RoboDK station: reto.rdk

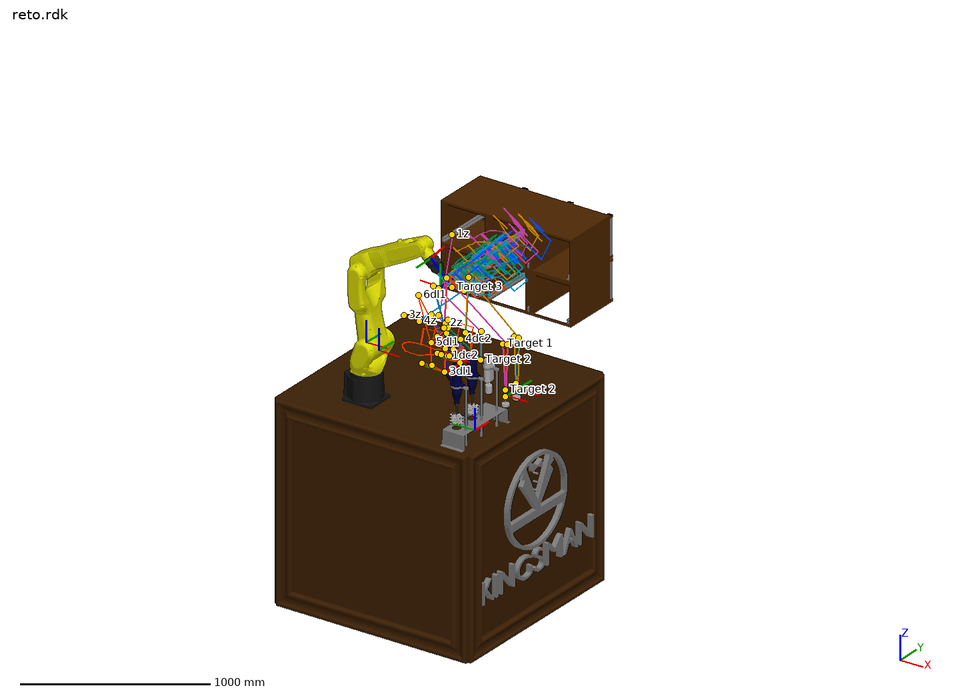
[picture v0: the station drawn from its stored meshes, robots at their saved joint values, targets as dots, program paths as lines]
Station reto (saved by RoboDK 5.5.4). Poses are relative to the parent item; angles as X-Y-Z fixed-axis rotations.
  - frame Fanuc LR Mate 200iD/7L Base at (0, 670, 330) mm
    - robot Fanuc LR Mate 200iD/7L: 6 axes, payload 7 kg, reach 911 mm, repeatability 0.03 mm, weight 27 kg
        modified DH rows (alpha deg, a mm, theta deg, d mm): 0, 0, 0, 330; -90, 50, -90, 0; 0, 440, 0, 0; -90, 35, 0, 420; 90, 0, 0, 0; -90, 0, 0, 80
        base shift (0, 0, -330) mm
        joint limits [-170, -70, -70, -190, -115, -360] to [170, 145, 215, 190, 115, 360]; home [0, 0, 0, 0, 0, 0]; saved at [0, -7.035, 27.253, 0, -70.54, 0]
      - frame RobotiQ 2F-140 Gripper (Mechanism) Base at (0, 0, 0) mm
        - robot RobotiQ 2F-140 Gripper (Mechanism) (model RobotiQ 2F140): 1 axes, payload 5 kg
            joint limits [0] to [140]; home [140]; saved at [30]
          - tool Tool 1, TCP at (0, 0, 190) mm
        - target open (joint target) at (-0.21, -35.16, 190) mm, rotated rx 0 ry -3.02 rz -0.35 deg; joints [30] of RobotiQ 2F-140 Gripper (Mechanism)
        - target close (joint target) at (-114.65, -295.92, 10.81) mm, rotated rx -1.72 ry 2.03 rz 11.69 deg; joints [10] of RobotiQ 2F-140 Gripper (Mechanism)
        - target Target 3 (Cartesian target) at (0, 0, 190) mm; joints [23.986, 137.128, 3.759, 0, 86.241, -156.014] of Fanuc LR Mate 200iD/7L
        - target Target 4 (Cartesian target) at (0, 0, 190) mm; joints [23.986, 137.128, 3.759, 0, 86.241, -156.014] of Fanuc LR Mate 200iD/7L
    - target home (Cartesian target) at (550, 0, 475) mm, rotated rx -180 ry -46.71 rz 0 deg; joints [0, 3.939, 7.691, 0, -50.978, 0] of Fanuc LR Mate 200iD/7L
  - frame rack at (-170, 1590, 240) mm, rotated rx 90 ry 0 rz 180 deg
    - object FullRack (1) at (-810, 360, -320) mm, size 835 x 510 x 385.3 mm, geometry from FullRack (1).STEP
    - target 1z (Cartesian target) at (-358.1, 564.97, -403.2) mm, rotated rx -26.57 ry -40.12 rz 107.86 deg; joints [70, -7.04, 27.25, 0, -70.54, 0] of Fanuc LR Mate 200iD/7L
    - target 2z (Cartesian target) at (-342.39, 58.73, -444.89) mm, rotated rx 2.43 ry -28.49 rz 101.39 deg; joints [48.708, 3.516, -60.085, -111.282, -47, 134.319] of Fanuc LR Mate 200iD/7L
    - target 3z (Cartesian target) at (-104.58, 56.68, -482.72) mm, rotated rx 2.43 ry -28.49 rz 101.39 deg; joints [97.474, -14.415, -55.536, -177.531, -28.246, 164.28] of Fanuc LR Mate 200iD/7L
    - target 4z (Cartesian target) at (-165.76, 16.78, -430.34) mm, rotated rx 2.43 ry -28.49 rz 101.39 deg; joints [82.687, 5.107, -71.647, -159.69, -45.234, 158.787] of Fanuc LR Mate 200iD/7L
    - target 5z (Cartesian target) at (-150, 20, 0) mm, rotated rx 2.43 ry -28.49 rz 101.39 deg; joints [88.603, 43.78, -43.517, 30.239, 18.18, -38.415] of Fanuc LR Mate 200iD/7L
    - target subida charola (Cartesian target) at (-343.88, 69.1, -423.53) mm, rotated rx -21.12 ry -28.57 rz 104.68 deg; joints [68.168, -3.801, -53.905, 12.841, 22.763, -13.527] of Fanuc LR Mate 200iD/7L
  - frame base herramental at (710, 650, 20) mm, rotated rx 0 ry 0 rz 90 deg
    - object Soporte de herramientas at (0, 0, 70) mm, rotated rx 90 ry 0 rz 180 deg, size 443.6 x 340 x 140 mm, geometry from Soporte de herramientas.STEP
  - frame dremel2 at (620, 650, 390) mm, rotated rx 0 ry 0 rz 90 deg
    - target 1dc2 (Cartesian target) at (0.49, 88.9, 17.55) mm, rotated rx -180 ry -61.75 rz -90 deg; joints [89.913, -3.297, -48.984, 180.078, 102.766, 0.058] of Fanuc LR Mate 200iD/7L
    - target 2dc2 (Cartesian target) at (0, 151.76, 13.3) mm, rotated rx -180 ry -61.75 rz -90 deg; joints [-4.961, -25.961, -32.248, 48.26, 5.86, -45.758] of Fanuc LR Mate 200iD/7L
    - target 3dc2 (Cartesian target) at (0, 4.92, 1.2) mm, rotated rx -180 ry -49.6 rz -90 deg; joints [-2.796, -1.172, -33.671, 162.466, 7.084, -160.778] of Fanuc LR Mate 200iD/7L
    - target 4dc2 (Cartesian target) at (0, 0.76, 138.38) mm, rotated rx -180 ry -49.6 rz -90 deg; joints [-2.768, -6.859, -13.429, 175.365, 27.075, -174.076] of Fanuc LR Mate 200iD/7L
    - target 5dc2 (Cartesian target) at (0, 92.68, 148.84) mm, rotated rx -180 ry -44.51 rz -90 deg; joints [-3.386, -17.516, -7.24, 176.175, 38.363, -174.583] of Fanuc LR Mate 200iD/7L
    - target 6dc2 (Cartesian target) at (477.83, 510, 116.81) mm, rotated rx -180 ry -49.6 rz 3.55 deg; joints [64.081, -25.306, -11.026, 143.659, 39.225, -130.203] of Fanuc LR Mate 200iD/7L
  - frame dremel1 at (620, 510.31, 389.97) mm, rotated rx 0 ry 0 rz 90 deg
    - target 1dl1 (Cartesian target) at (0.49, 88.9, 17.55) mm, rotated rx -180 ry -61.75 rz -90 deg; joints [-28.495, -9.165, -37.687, 76.78, 25.575, -60.993] of Fanuc LR Mate 200iD/7L
    - target 2dl1 (Cartesian target) at (0, 151.76, 13.3) mm, rotated rx -180 ry -61.75 rz -90 deg; joints [-34.725, -17.114, -36.143, 84.899, 30.251, -65.939] of Fanuc LR Mate 200iD/7L
    - target 3dl1 (Cartesian target) at (0, 4.92, 1.2) mm, rotated rx -180 ry -49.6 rz -90 deg; joints [-21.306, 2.651, -33.616, 117.955, 18.257, -105.014] of Fanuc LR Mate 200iD/7L
    - target 4dl1 (Cartesian target) at (0, 0.76, 138.38) mm, rotated rx -180 ry -48.03 rz -90 deg; joints [-20.886, -2.493, -13.042, 151.816, 34.141, -141.769] of Fanuc LR Mate 200iD/7L
    - target 5dl1 (Cartesian target) at (0, 92.68, 148.84) mm, rotated rx -180 ry -49.6 rz -90 deg; joints [-26.4, -14.504, -10.508, 146.56, 37.916, -134.648] of Fanuc LR Mate 200iD/7L
    - target 6dl1 (Cartesian target) at (477.83, 510, 116.81) mm, rotated rx -180 ry -55.33 rz 3.55 deg; joints [37.94, -45.517, -1.764, 129.234, 61.201, -109.727] of Fanuc LR Mate 200iD/7L
    - object cepillo1 at (0, -70, -50) mm, rotated rx 90 ry 0 rz 180 deg, size 80 x 351.1 x 124.1 mm, geometry from Dremel con brida.STEP
  - frame bote cera at (140, 586, 355) mm
    - target Target 1 (Cartesian target) at (316.19, 84, 136.54) mm, rotated rx -180 ry -46.71 rz 0 deg; joints [0, -28.492, -10.215, 0, -33.072, 0] of Fanuc LR Mate 200iD/7L
    - target Target 3 (Cartesian target) at (300.65, 202.07, 136.5) mm, rotated rx -180 ry -46.9 rz 15 deg; joints [15, -28.576, -10.266, 0, -32.834, 0] of Fanuc LR Mate 200iD/7L
    - target Target 2 (Cartesian target) at (513.63, 198.92, 10) mm, rotated rx -180 ry -50.56 rz 10.82 deg; joints [9.584, 6.819, -37.897, -31.652, -1.82, 32.424] of Fanuc LR Mate 200iD/7L
    - target Target 4 (Cartesian target) at (516.39, 196.06, 177.59) mm, rotated rx -179.95 ry -49.71 rz 10.96 deg; joints [9.091, -0.877, -13.325, -3.243, -27.022, 4.097] of Fanuc LR Mate 200iD/7L
    - target Target 5 (Cartesian target) at (-35.2, 592.88, 112.91) mm, rotated rx 179.59 ry -46.7 rz 80 deg; joints [77.715, -18.214, -17.774, -2.891, -25.565, 4.172] of Fanuc LR Mate 200iD/7L
  - program open (3 instructions, listed below)
  - program close (3 instructions, listed below)
  - program home (4 instructions, listed below)
  - object mesa at (-1220, 1130, 330) mm, size 1277.5 x 1274.9 x 1205 mm, geometry from mesa.STEP
  - frame zapato at (110, 1270, 40) mm
    - target Target 1 (Cartesian target) at (78.1, -83.2, 764.97) mm, rotated rx -180 ry -46.71 rz 70 deg; joints [70, -7.04, 27.25, 0, -70.54, 0] of Fanuc LR Mate 200iD/7L
    - target Target 2 (Cartesian target) at (48.8, -163.69, 316.74) mm, rotated rx -179.51 ry -45.09 rz 70 deg; joints [69.514, -19.906, -32.534, -3.891, -12.407, 4.144] of Fanuc LR Mate 200iD/7L
    - target Target 3 (Cartesian target) at (51.99, -36.78, 68.56) mm, rotated rx -167.65 ry -61.99 rz 84.86 deg; joints [58.654, 42.845, -90.321, 40.028, 62.94, -6.257] of Fanuc LR Mate 200iD/7L
    - target Target 4 (Cartesian target) at (0, 0, 0) mm, rotated rx -154.66 ry -59.5 rz 70 deg; joints [67.996, 54.587, -97.1, 29.193, 68.847, -10.257] of Fanuc LR Mate 200iD/7L
    - target Target 5 (Cartesian target) at (-12.96, -146.91, 298.71) mm, rotated rx -168.48 ry -59.46 rz 67.92 deg; joints [74.53, -18.6, -45.29, -158.86, -16.3, 156.27] of Fanuc LR Mate 200iD/7L
    - target Target 6 (Cartesian target) at (14.48, -93.65, 48.92) mm, rotated rx -154.66 ry -59.5 rz 70 deg; joints [59.102, 46.97, -102.654, -143.53, -72.674, 174.279] of Fanuc LR Mate 200iD/7L
  - program recoger cepillo cera (10 instructions, listed below)
  - program reset (1 instructions, listed below)
  - program recoger cepillo limpieza (10 instructions, listed below)
  - program recoger cera (9 instructions, listed below)
  - program pick charola (8 instructions, listed below)
  - program c1 recoger (7 instructions, listed below)
  - program c1 entregar (7 instructions, listed below)
  - program poscharolamesa (7 instructions, listed below)
  - program dejar cepillo limpieza (9 instructions, listed below)
  - program dejar cepillo cera (10 instructions, listed below)
  - program dejar  cera (9 instructions, listed below)
  - machining project parribaizq: rotZ(0) | rotX(0)*rotY(0) | onStart | onPathStart | onApproach | onPoint | onRetract | onFinish | SetRPM(%1) | SetTool(%1) | Extruder(%1) | default | default | OutOnMov(%1) | OutOffMov(%1) | onPathFinish | M_RunCode(%1)
  - machining project plateralesizq: rotZ(0) | rotX(0)*rotY(0) | onStart | onPathStart | onApproach | onPoint | onRetract | onFinish | SetRPM(%1) | SetTool(%1) | Extruder(%1) | default | default | OutOnMov(%1) | OutOffMov(%1) | onPathFinish | M_RunCode(%1)
  - program parrizq (66 instructions, listed below)
  - machining project Path3 ajustes: rotZ(0) | rotX(0)*rotY(0) | onStart | onPathStart | onApproach | onPoint | onRetract | onFinish | SetRPM(%1) | SetTool(%1) | Extruder(%1) | default | default | OutOnMov(%1) | OutOffMov(%1) | onPathFinish | M_RunCode(%1)
  - machining project Path4 ajustes: rotZ(0) | rotX(0)*rotY(0) | onStart | onPathStart | onApproach | onPoint | onRetract | onFinish | SetRPM(%1) | SetTool(%1) | Extruder(%1) | default | default | OutOnMov(%1) | OutOffMov(%1) | onPathFinish | M_RunCode(%1)
  - program parrder (59 instructions, listed below)
  - program final (30 instructions, listed below)
  - machining project Path5 ajustes: rotZ(0) | rotX(0)*rotY(0) | onStart | onPathStart | onApproach | onPoint | onRetract | onFinish | SetRPM(%1) | SetTool(%1) | Extruder(%1) | default | default | OutOnMov(%1) | OutOffMov(%1) | onPathFinish | M_RunCode(%1)
  - program cerlatizq (163 instructions, listed below)
  - program platder (154 instructions, listed below)
  - machining project Path6 ajustes: rotZ(0) | rotX(0)*rotY(0) | onStart | onPathStart | onApproach | onPoint | onRetract | onFinish | SetRPM(%1) | SetTool(%1) | Extruder(%1) | default | default | OutOnMov(%1) | OutOffMov(%1) | onPathFinish | M_RunCode(%1)
  - program platizq (163 instructions, listed below)
  - program carribizq (66 instructions, listed below)
  - machining project Path7 ajustes: rotZ(0) | rotX(0)*rotY(0) | onStart | onPathStart | onApproach | onPoint | onRetract | onFinish | SetRPM(%1) | SetTool(%1) | Extruder(%1) | default | default | OutOnMov(%1) | OutOffMov(%1) | onPathFinish | M_RunCode(%1)
  - program cerlatder (154 instructions, listed below)
  - machining project Path8 ajustes: rotZ(0) | rotX(0)*rotY(0) | onStart | onPathStart | onApproach | onPoint | onRetract | onFinish | SetRPM(%1) | SetTool(%1) | Extruder(%1) | default | default | OutOnMov(%1) | OutOffMov(%1) | onPathFinish | M_RunCode(%1)
  - program cerarribder (44 instructions, listed below)
  - machining project Path10 ajustes: rotZ(0) | rotX(0)*rotY(0) | onStart | onPathStart | onApproach | onPoint | onRetract | onFinish | SetRPM(%1) | SetTool(%1) | Extruder(%1) | default | default | OutOnMov(%1) | OutOffMov(%1) | onPathFinish | M_RunCode(%1)
  - program talonder (20 instructions, listed below)
  - frame iman izquierdo at (690, 970, 90) mm, rotated rx 0 ry -0.43 rz 0 deg
    - target Target 1 (Cartesian target) at (-16, -10, 304.12) mm, rotated rx -180 ry -3.01 rz 0 deg; joints [23.726, 34.659, -8.597, 1.235, -78.648, -23.94] of Fanuc LR Mate 200iD/7L
    - target Target 2 (Cartesian target) at (-1.94, -10, 36.88) mm, rotated rx -180 ry -3.01 rz 0 deg; joints [23.284, 48.242, -37.276, 1.554, -49.968, -24.255] of Fanuc LR Mate 200iD/7L
    - target Target 3 (Cartesian target) at (-0.39, -10, 0.32) mm, rotated rx -180 ry 2.75 rz 0 deg; joints [22.488, 53.778, -37.823, -1.092, -54.324, -21.835] of Fanuc LR Mate 200iD/7L
    - target Target 4 (Cartesian target) at (14.23, -10, 304.96) mm, rotated rx -180 ry 2.75 rz 0 deg; joints [22.137, 42.684, -3.214, -0.874, -88.934, -22.104] of Fanuc LR Mate 200iD/7L
    - target Target 5 (Cartesian target) at (-604.68, 318.92, 397.91) mm, rotated rx -178.71 ry 2.21 rz 80.14 deg; joints [82.014, 21.757, -2.792, -0.939, -89.319, -1.878] of Fanuc LR Mate 200iD/7L
    - target Target 6 (Cartesian target) at (-653.05, 360.19, 74.8) mm, rotated rx -178.71 ry 0.13 rz 80.09 deg; joints [86.488, 37.843, -40.739, -1.149, -49.231, -5.645] of Fanuc LR Mate 200iD/7L
  - frame iman derecho at (690, 1070, 90) mm
    - target Target 1 (Cartesian target) at (-16, -10, 304.12) mm, rotated rx -180 ry -3.01 rz 0 deg; joints [30.586, 42.114, -3.765, 1.541, -83.645, -30.722] of Fanuc LR Mate 200iD/7L
    - target Target 2 (Cartesian target) at (-1.94, -10, 36.88) mm, rotated rx -180 ry -3.01 rz 0 deg; joints [30.06, 53.677, -32.189, 1.836, -55.219, -31.073] of Fanuc LR Mate 200iD/7L
    - target Target 3 (Cartesian target) at (-0.39, -0.58, 0.32) mm, rotated rx -180 ry 2.75 rz 0 deg; joints [29.619, 60.126, -31.432, -1.553, -60.966, -28.837] of Fanuc LR Mate 200iD/7L
    - target Target 4 (Cartesian target) at (14.23, -10, 304.96) mm, rotated rx -180 ry 2.75 rz 0 deg; joints [28.537, 52.814, 4.62, -1.322, -97.032, -28.672] of Fanuc LR Mate 200iD/7L
    - target Target 5 (Cartesian target) at (-491.92, 250.35, 416.93) mm, rotated rx -178.68 ry 2.41 rz 72.7 deg; joints [72.54, 30.81, 4.62, -1.32, -97.03, 0] of Fanuc LR Mate 200iD/7L
    - target Target 6 (Cartesian target) at (-525.43, 271.58, 73.13) mm, rotated rx -178.86 ry -1.69 rz 77.54 deg; joints [75.764, 40.036, -38.477, -1.565, -49.877, 2.787] of Fanuc LR Mate 200iD/7L
  - program iman izquierdo (13 instructions, listed below)
  - program iman derecho (13 instructions, listed below)
  - program dejar iman izquierdo (12 instructions, listed below)
  - program dejar iman derecho (12 instructions, listed below)
  - machining project Path10 ajustes: rotZ(0) | rotX(0)*rotY(0) | onStart | onPathStart | onApproach | onPoint | onRetract | onFinish | SetRPM(%1) | SetTool(%1) | Extruder(%1) | default | default | OutOnMov(%1) | OutOffMov(%1) | onPathFinish | M_RunCode(%1)
  - program platizch (163 instructions, listed below)
  - machining project Path11 ajustes: rotZ(0) | rotX(0)*rotY(0) | onStart | onPathStart | onApproach | onPoint | onRetract | onFinish | SetRPM(%1) | SetTool(%1) | Extruder(%1) | default | default | OutOnMov(%1) | OutOffMov(%1) | onPathFinish | M_RunCode(%1)
  - program plaizgr (163 instructions, listed below)
  - machining project Path12 ajustes: rotZ(0) | rotX(0)*rotY(0) | onStart | onPathStart | onApproach | onPoint | onRetract | onFinish | SetRPM(%1) | SetTool(%1) | Extruder(%1) | default | default | OutOnMov(%1) | OutOffMov(%1) | onPathFinish | M_RunCode(%1)
  - program pladerch (154 instructions, listed below)
  - machining project Path13 ajustes: rotZ(0) | rotX(0)*rotY(0) | onStart | onPathStart | onApproach | onPoint | onRetract | onFinish | SetRPM(%1) | SetTool(%1) | Extruder(%1) | default | default | OutOnMov(%1) | OutOffMov(%1) | onPathFinish | M_RunCode(%1)
  - program pladergr (154 instructions, listed below)
  - machining project Path14 ajustes: rotZ(0) | rotX(0)*rotY(0) | onStart | onPathStart | onApproach | onPoint | onRetract | onFinish | SetRPM(%1) | SetTool(%1) | Extruder(%1) | default | default | OutOnMov(%1) | OutOffMov(%1) | onPathFinish | M_RunCode(%1)
  - program arrizch (57 instructions, listed below)
  - machining project Path15 ajustes: rotZ(0) | rotX(0)*rotY(0) | onStart | onPathStart | onApproach | onPoint | onRetract | onFinish | SetRPM(%1) | SetTool(%1) | Extruder(%1) | default | default | OutOnMov(%1) | OutOffMov(%1) | onPathFinish | M_RunCode(%1)
  - program arriderch (52 instructions, listed below)
  - machining project Path16 ajustes: rotZ(0) | rotX(0)*rotY(0) | onStart | onPathStart | onApproach | onPoint | onRetract | onFinish | SetRPM(%1) | SetTool(%1) | Extruder(%1) | default | default | OutOnMov(%1) | OutOffMov(%1) | onPathFinish | M_RunCode(%1)
  - program arridergr (59 instructions, listed below)
  - machining project Path17 ajustes: rotZ(0) | rotX(0)*rotY(0) | onStart | onPathStart | onApproach | onPoint | onRetract | onFinish | SetRPM(%1) | SetTool(%1) | Extruder(%1) | default | default | OutOnMov(%1) | OutOffMov(%1) | onPathFinish | M_RunCode(%1)
  - program arriizqgr (57 instructions, listed below)
  - machining project Path18 ajustes: rotZ(0) | rotX(0)*rotY(0) | onStart | onPathStart | onApproach | onPoint | onRetract | onFinish | SetRPM(%1) | SetTool(%1) | Extruder(%1) | default | default | OutOnMov(%1) | OutOffMov(%1) | onPathFinish | M_RunCode(%1)
  - program cerlaizgr (163 instructions, listed below)
  - machining project Path19 ajustes: rotZ(0) | rotX(0)*rotY(0) | onStart | onPathStart | onApproach | onPoint | onRetract | onFinish | SetRPM(%1) | SetTool(%1) | Extruder(%1) | default | default | OutOnMov(%1) | OutOffMov(%1) | onPathFinish | M_RunCode(%1)
  - program cerladergr (154 instructions, listed below)
  - machining project Path20 ajustes: rotZ(0) | rotX(0)*rotY(0) | onStart | onPathStart | onApproach | onPoint | onRetract | onFinish | SetRPM(%1) | SetTool(%1) | Extruder(%1) | default | default | OutOnMov(%1) | OutOffMov(%1) | onPathFinish | M_RunCode(%1)
  - program ceraariizgr (59 instructions, listed below)
  - machining project Path21 ajustes: rotZ(0) | rotX(0)*rotY(0) | onStart | onPathStart | onApproach | onPoint | onRetract | onFinish | SetRPM(%1) | SetTool(%1) | Extruder(%1) | default | default | OutOnMov(%1) | OutOffMov(%1) | onPathFinish | M_RunCode(%1)
  - program cerarridergr (59 instructions, listed below)
  - machining project Path22 ajustes: rotZ(0) | rotX(0)*rotY(0) | onStart | onPathStart | onApproach | onPoint | onRetract | onFinish | SetRPM(%1) | SetTool(%1) | Extruder(%1) | default | default | OutOnMov(%1) | OutOffMov(%1) | onPathFinish | M_RunCode(%1)
  - program cerlatizqch (163 instructions, listed below)
  - machining project Path23 ajustes: rotZ(0) | rotX(0)*rotY(0) | onStart | onPathStart | onApproach | onPoint | onRetract | onFinish | SetRPM(%1) | SetTool(%1) | Extruder(%1) | default | default | OutOnMov(%1) | OutOffMov(%1) | onPathFinish | M_RunCode(%1)
  - program cerlatderch (154 instructions, listed below)
  - machining project Path25 ajustes: rotZ(0) | rotX(0)*rotY(0) | onStart | onPathStart | onApproach | onPoint | onRetract | onFinish | SetRPM(%1) | SetTool(%1) | Extruder(%1) | default | default | OutOnMov(%1) | OutOffMov(%1) | onPathFinish | M_RunCode(%1)
  - program ceraarribderch (59 instructions, listed below)
  - machining project Path26 ajustes: rotZ(0) | rotX(0)*rotY(0) | onStart | onPathStart | onApproach | onPoint | onRetract | onFinish | SetRPM(%1) | SetTool(%1) | Extruder(%1) | default | default | OutOnMov(%1) | OutOffMov(%1) | onPathFinish | M_RunCode(%1)
  - program ceraarribaizqch (59 instructions, listed below)
  - program final_ch (30 instructions, listed below)
  - program final_gr (30 instructions, listed below)
  - object cepillo2 at (690, 650, 340) mm, rotated rx 90 ry 0 rz -90 deg, size 80 x 351.1 x 124.1 mm, geometry from Dremel con brida.STEP
  - object Iman at (688.21, 960, 126.59) mm, rotated rx 90 ry 0 rz 0 deg, size 45.7 x 91.4 x 45.7 mm, geometry from Iman.STEP
  - object Iman at (688.48, 1060.58, 126.61) mm, size 45.7 x 91.4 x 45.7 mm, geometry from Iman.STEP
  - object Grasa  at (650, 792, 370) mm, size 75 x 201.5 x 85 mm, geometry from Grasa (1).STEP
  - object zapatoconcharola at (-21.13, 1591.46, 262.04) mm, rotated rx 0 ry 0 rz -0.01 deg, size 250 x 350 x 100.5 mm, geometry from zapatoconcharola.STEP
    - object Ruta_IZQ at (-60, 470, 60) mm, rotated rx 0 ry 0 rz -90 deg, geometry from Curva importada
    - object R7 at (-105, 460, 60) mm, rotated rx 0 ry 0 rz -90 deg
    - object Ruta_IZQ_ch at (-60, 390, 60) mm, rotated rx 0 ry 0 rz -90 deg, geometry from Curva importada
    - object R7_ch at (-67.5, 380, 60) mm, rotated rx 0 ry 0 rz -90 deg
    - object Ruta_IZQ_gr at (-50, 550, 80) mm, rotated rx 0 ry 0 rz -90 deg, geometry from Curva importada
    - object R7_gr at (-135, 550, 80) mm, rotated rx 0 ry 0 rz -90 deg
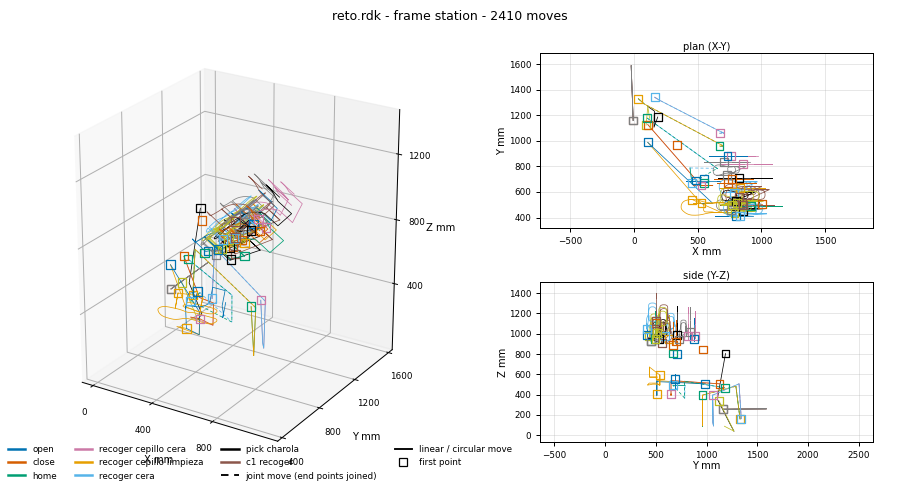
[picture p0: tool path of reto.rdk in frame station, 2410 of 2410 moves have a stored position in this frame; points joined in program order, loops and branches not executed]

--- program open (robot RobotiQ 2F-140 Gripper (Mechanism)) ---
  Est. Ref.: RobotiQ 2F-140 Gripper (Mechanism) Base
  Est. herr: Tool 1
  MoveJ (open)

--- program close (robot RobotiQ 2F-140 Gripper (Mechanism)) ---
  Est. Ref.: RobotiQ 2F-140 Gripper (Mechanism) Base
  Est. herr: Tool 1
  MoveJ (close)

--- program home (robot Fanuc LR Mate 200iD/7L) ---
  Est. Ref.: Fanuc LR Mate 200iD/7L Base
  MoveJ (home)
  Llamar open
  Separar de Tool 1

--- program recoger cepillo cera (robot Fanuc LR Mate 200iD/7L) ---
  Est. Ref.: dremel2
  Est. herr: Tool 1
  MoveL (1dc2)
  MoveL (Target 2) -> target 2dc2
  MoveL (Target 3) -> target 3dc2
  Llamar close
  Adjuntar a Tool 1
  MoveL (Target 4) -> target 4dc2
  MoveL (Target 5) -> target 5dc2
  MoveL (6dc2)

--- program reset (robot Fanuc LR Mate 200iD/7L) ---
  Reemplazar objetos

--- program recoger cepillo limpieza (robot Fanuc LR Mate 200iD/7L) ---
  Est. Ref.: dremel1
  Est. herr: Tool 1
  MoveL (1dl1)
  MoveL (2dl1)
  MoveL (3dl1)
  Adjuntar a Tool 1
  Llamar close
  MoveL (4dl1)
  MoveL (5dl1)
  MoveL (6dl1)

--- program recoger cera (robot Fanuc LR Mate 200iD/7L) ---
  Est. Ref.: bote cera
  Est. herr: Tool 1
  MoveJ (Target 1)
  MoveL (Target 3)
  MoveJ (Target 2)
  Llamar close
  Adjuntar a Tool 1
  MoveJ (Target 4)
  MoveL (Target 5)

--- program pick charola (robot Fanuc LR Mate 200iD/7L) ---
  Est. Ref.: zapato
  Est. herr: Tool 1
  MoveJ (Target 1)
  MoveL (Target 2)
  MoveL (Target 3)
  MoveL (Target 4)
  Llamar close
  Adjuntar a Tool 1

--- program c1 recoger (robot Fanuc LR Mate 200iD/7L) ---
  Est. Ref.: rack
  Est. herr: Tool 1
  MoveL (4z)
  MoveL (Target 4) -> target 5z
  Adjuntar a Tool 1
  Llamar close
  MoveL (4z)

--- program c1 entregar (robot Fanuc LR Mate 200iD/7L) ---
  Est. Ref.: rack
  Est. herr: Tool 1
  MoveL (4z)
  MoveL (Target 4) -> target 5z
  Separar de Tool 1
  Llamar open
  MoveL (4z)

--- program poscharolamesa (robot Fanuc LR Mate 200iD/7L) ---
  Est. Ref.: zapato
  Est. herr: Tool 1
  MoveJ (Target 5)
  MoveL (Target 4)
  Separar de Tool 1
  Llamar open
  MoveL (Target 6)

--- program dejar cepillo limpieza (robot Fanuc LR Mate 200iD/7L) ---
  Est. Ref.: dremel1
  Est. herr: Tool 1
  MoveL (6dl1)
  MoveL (4dl1)
  MoveL (3dl1)
  Separar de Tool 1
  Llamar open
  MoveL (1dl1)
  MoveL (5dl1)

--- program dejar cepillo cera (robot Fanuc LR Mate 200iD/7L) ---
  Est. Ref.: dremel2
  Est. herr: Tool 1
  MoveL (6dc2)
  MoveL (Target 5) -> target 5dc2
  MoveL (Target 4) -> target 4dc2
  MoveL (Target 3) -> target 3dc2
  Llamar open
  Separar de Tool 1
  MoveL (1dc2)
  MoveL (Target 2) -> target 2dc2

--- program dejar  cera (robot Fanuc LR Mate 200iD/7L) ---
  Est. Ref.: bote cera
  Est. herr: Tool 1
  MoveL (Target 5)
  MoveJ (Target 4)
  MoveJ (Target 2)
  Llamar open
  Separar de Tool 1
  MoveJ (Target 1)
  MoveL (Target 3)

--- program parrizq (robot Fanuc LR Mate 200iD/7L) ---
  Suave(1)
  Establecer velocidad (1000.0 mm/s)
  Est. Ref.: RobotiQ 2F-140 Gripper (Mechanism) Base
  Est. herr: Tool 1
  Mostrar Tool 1
  MoveJ 1 to (272.96, -213.5, 226.79) mm, rotated rx 167 ry 29.36 rz -96.45 deg; joints [111.702, 50.919, -11.475, 32.192, -81.814, 59.615]
  MoveL 2 to (272.96, -213.5, 226.79) mm, rotated rx 167 ry 29.36 rz -96.45 deg; joints [111.702, 50.919, -11.475, 32.192, -81.814, 59.615]
  MoveL 3 to (253.35, -213.5, 128.73) mm, rotated rx 167 ry 29.36 rz -96.45 deg; joints [111.201, 57.407, -19.462, 33.135, -74.825, 55.631]
  MoveL 4 to (253.35, -213.5, 128.73) mm, rotated rx 167 ry 29.36 rz -96.45 deg; joints [111.201, 57.407, -19.462, 33.135, -74.825, 55.631]
  Establecer velocidad (50.0 mm/s)
  MoveL 5 to (243.62, -213.5, 127.58) mm, rotated rx 167 ry 29.36 rz -96.45 deg; joints [110.96, 59.057, -18.114, 32.97, -75.831, 56.589]
  MoveL 6 to (233.9, -213.5, 126.22) mm, rotated rx 167 ry 29.36 rz -96.45 deg; joints [110.725, 60.817, -16.674, 32.805, -76.918, 57.588]
  MoveL 7 to (223.13, -213.5, 124.47) mm, rotated rx 167 ry 29.36 rz -96.45 deg; joints [110.47, 62.925, -14.939, 32.622, -78.246, 58.759]
  MoveL 8 to (210.98, -213.5, 122.18) mm, rotated rx 167 ry 29.36 rz -96.45 deg; joints [110.189, 65.575, -12.731, 32.417, -79.961, 60.202]
  MoveL 9 to (200.56, -213.5, 119.96) mm, rotated rx 167 ry 29.36 rz -96.45 deg; joints [109.954, 68.174, -10.522, 32.242, -81.705, 61.595]
  MoveL 10 to (195.63, -213.5, 118.82) mm, rotated rx 167 ry 29.36 rz -96.45 deg; joints [109.845, 69.562, -9.321, 32.16, -82.664, 62.333]
  MoveL 11 to (191.25, -213.5, 117.76) mm, rotated rx 167 ry 29.36 rz -96.45 deg; joints [109.749, 70.916, -8.132, 32.089, -83.62, 63.051]
  MoveL 12 to (189.42, -213.5, 117.22) mm, rotated rx 167 ry 29.36 rz -96.45 deg; joints [109.709, 71.53, -7.597, 32.06, -84.052, 63.371]
  MoveL 13 to (188.23, -213.5, 116.45) mm, rotated rx 167 ry 29.36 rz -96.45 deg; joints [109.683, 71.949, -7.286, 32.045, -84.302, 63.558]
  MoveL 14 to (187.22, -213.5, 115.14) mm, rotated rx 167 ry 29.36 rz -96.45 deg; joints [109.661, 72.325, -7.09, 32.035, -84.457, 63.681]
  MoveL 15 to (186.8, -213.5, 113.88) mm, rotated rx 167 ry 29.36 rz -96.45 deg; joints [109.652, 72.499, -7.088, 32.036, -84.453, 63.69]
  MoveL 16 to (186.72, -213.5, 112.35) mm, rotated rx 167 ry 29.36 rz -96.45 deg; joints [109.65, 72.551, -7.244, 32.044, -84.32, 63.608]
  MoveL 17 to (186.72, -213.5, 110.28) mm, rotated rx 167 ry 29.36 rz -96.45 deg; joints [109.65, 72.587, -7.49, 32.057, -84.112, 63.477]
  MoveL 18 to (186.72, -213.5, 106.61) mm, rotated rx 167 ry 29.36 rz -96.45 deg; joints [109.65, 72.658, -7.92, 32.081, -83.748, 63.248]
  MoveL 19 to (186.72, -213.5, 102.35) mm, rotated rx 167 ry 29.36 rz -96.45 deg; joints [109.65, 72.751, -8.407, 32.111, -83.335, 62.987]
  MoveL 20 to (186.72, -213.5, 98.08) mm, rotated rx 167 ry 29.36 rz -96.45 deg; joints [109.65, 72.855, -8.884, 32.141, -82.931, 62.732]
  MoveL 21 to (186.72, -213.5, 93.7) mm, rotated rx 167 ry 29.36 rz -96.45 deg; joints [109.65, 72.974, -9.362, 32.174, -82.526, 62.475]
  Establecer velocidad (1000.0 mm/s)
  MoveL 22 to (186.72, -213.5, 93.7) mm, rotated rx 167 ry 29.36 rz -96.45 deg; joints [109.65, 72.974, -9.362, 32.174, -82.526, 62.475]
  MoveL 23 to (206.33, -213.5, 191.76) mm, rotated rx 167 ry 29.36 rz -96.45 deg; joints [110.083, 65.723, -3.105, 31.883, -88.061, 65.437]
  Establecer velocidad (1000.0 mm/s)
  MoveL 24 to (282.76, -213.5, 227.74) mm, rotated rx 167 ry 29.36 rz -96.45 deg; joints [111.961, 49.296, -12.655, 32.266, -80.951, 58.762]
  MoveL 25 to (263.15, -213.5, 129.69) mm, rotated rx 167 ry 29.36 rz -96.45 deg; joints [111.449, 55.838, -20.746, 33.301, -73.879, 54.698]
  MoveL 26 to (263.15, -213.5, 129.69) mm, rotated rx 167 ry 29.36 rz -96.45 deg; joints [111.449, 55.838, -20.746, 33.301, -73.879, 54.698]
  Establecer velocidad (50.0 mm/s)
  MoveL 27 to (281.65, -213.5, 132.2) mm, rotated rx 167 ry 29.36 rz -96.45 deg; joints [111.932, 53.024, -22.888, 33.594, -72.339, 53.073]
  MoveL 28 to (301.97, -213.5, 137.15) mm, rotated rx 167 ry 29.36 rz -96.45 deg; joints [112.488, 50.029, -24.766, 33.854, -71.059, 51.53]
  MoveL 29 to (321.64, -213.5, 144.29) mm, rotated rx 167 ry 29.36 rz -96.45 deg; joints [113.051, 47.158, -26.131, 34.028, -70.211, 50.275]
  MoveL 30 to (340.4, -213.5, 153.54) mm, rotated rx 167 ry 29.36 rz -96.45 deg; joints [113.614, 44.389, -27.009, 34.107, -69.766, 49.308]
  MoveL 31 to (358.05, -213.5, 164.78) mm, rotated rx 167 ry 29.36 rz -96.45 deg; joints [114.168, 41.717, -27.415, 34.089, -69.705, 48.63]
  MoveL 32 to (374.35, -213.5, 177.88) mm, rotated rx 167 ry 29.36 rz -96.45 deg; joints [114.702, 39.153, -27.366, 33.977, -70.011, 48.241]
  MoveL 33 to (389.14, -213.5, 192.68) mm, rotated rx 167 ry 29.36 rz -96.45 deg; joints [115.205, 36.717, -26.881, 33.784, -70.663, 48.133]
  Establecer velocidad (1000.0 mm/s)
  MoveL 34 to (389.14, -213.5, 192.68) mm, rotated rx 167 ry 29.36 rz -96.45 deg; joints [115.205, 36.717, -26.881, 33.784, -70.663, 48.133]
  MoveL 35 to (408.75, -213.5, 290.74) mm, rotated rx 167 ry 29.36 rz -96.45 deg; joints [115.902, 30.516, -16.673, 32.189, -79.585, 53.316]
  Establecer velocidad (1000.0 mm/s)
  MoveL 36 to (517.53, -213.5, 256.38) mm, rotated rx 167 ry 29.36 rz -96.45 deg; joints [120.525, 19.729, -26.554, 32.617, -73.54, 44.144]
  MoveL 37 to (497.92, -213.5, 158.32) mm, rotated rx 167 ry 29.36 rz -96.45 deg; joints [119.585, 27.601, -37.88, 35.349, -63.693, 38.061]
  MoveL 38 to (497.92, -213.5, 158.32) mm, rotated rx 167 ry 29.36 rz -96.45 deg; joints [119.585, 27.601, -37.88, 35.349, -63.693, 38.061]
  Establecer velocidad (50.0 mm/s)
  MoveL 39 to (500.24, -213.5, 142.39) mm, rotated rx 167 ry 29.36 rz -96.45 deg; joints [119.694, 28.554, -39.931, 35.928, -62.075, 36.641]
  MoveL 40 to (500.27, -213.5, 126.29) mm, rotated rx 167 ry 29.36 rz -96.45 deg; joints [119.695, 29.796, -41.859, 36.551, -60.522, 35.341]
  MoveL 41 to (498.03, -213.5, 110.35) mm, rotated rx 167 ry 29.36 rz -96.45 deg; joints [119.59, 31.286, -43.605, 37.197, -59.078, 34.2]
  MoveL 42 to (495.96, -213.5, 102.2) mm, rotated rx 167 ry 29.36 rz -96.45 deg; joints [119.494, 32.146, -44.426, 37.533, -58.384, 33.681]
  Establecer velocidad (1000.0 mm/s)
  MoveL 43 to (495.96, -213.5, 102.2) mm, rotated rx 167 ry 29.36 rz -96.45 deg; joints [119.494, 32.146, -44.426, 37.533, -58.384, 33.681]
  MoveL 44 to (515.57, -213.5, 200.26) mm, rotated rx 167 ry 29.36 rz -96.45 deg; joints [120.429, 23.061, -33.594, 34.007, -67.608, 40.119]
  Establecer velocidad (1000.0 mm/s)
  MoveL 45 to (517.53, -213.5, 256.38) mm, rotated rx 167 ry 29.36 rz -96.45 deg; joints [120.525, 19.729, -26.554, 32.617, -73.54, 44.144]
  MoveL 46 to (497.92, -213.5, 158.32) mm, rotated rx 167 ry 29.36 rz -96.45 deg; joints [119.585, 27.601, -37.88, 35.349, -63.693, 38.061]
  MoveL 47 to (497.92, -213.5, 158.32) mm, rotated rx 167 ry 29.36 rz -96.45 deg; joints [119.585, 27.601, -37.88, 35.349, -63.693, 38.061]
  Establecer velocidad (50.0 mm/s)
  MoveL 48 to (491.38, -213.5, 192.68) mm, rotated rx 167 ry 29.36 rz -96.45 deg; joints [119.283, 25.939, -33.348, 34.253, -67.275, 41.126]
  Establecer velocidad (1000.0 mm/s)
  MoveL 49 to (491.38, -213.5, 192.68) mm, rotated rx 167 ry 29.36 rz -96.45 deg; joints [119.283, 25.939, -33.348, 34.253, -67.275, 41.126]
  MoveL 50 to (510.99, -213.5, 290.74) mm, rotated rx 167 ry 29.36 rz -96.45 deg; joints [120.205, 18.932, -21.891, 32.036, -77.325, 46.974]

--- program parrder (robot Fanuc LR Mate 200iD/7L) ---
  Suave(1)
  Establecer velocidad (1000.0 mm/s)
  Est. Ref.: RobotiQ 2F-140 Gripper (Mechanism) Base
  Est. herr: Tool 1
  Mostrar Tool 1
  MoveJ 1 to (294.14, 36.7, 296.46) mm, rotated rx 168.69 ry 0 rz -89.99 deg; joints [86.744, 33.884, -9.121, -0.683, -69.59, 93.431]
  MoveL 2 to (294.14, 36.7, 296.46) mm, rotated rx 168.69 ry 0 rz -89.99 deg; joints [86.744, 33.884, -9.121, -0.683, -69.59, 93.431]
  MoveL 3 to (274.53, 36.7, 198.4) mm, rotated rx 168.69 ry 0 rz -89.99 deg; joints [86.831, 39.07, -19.388, -0.724, -59.322, 93.477]
  MoveL 4 to (274.53, 36.7, 198.4) mm, rotated rx 168.69 ry 0 rz -89.99 deg; joints [86.831, 39.07, -19.388, -0.724, -59.322, 93.477]
  Establecer velocidad (50.0 mm/s)
  MoveL 5 to (272.44, 36.7, 198.21) mm, rotated rx 168.69 ry 0 rz -89.99 deg; joints [86.84, 39.367, -19.213, -0.721, -59.497, 93.464]
  MoveL 6 to (270.34, 36.7, 198.02) mm, rotated rx 168.69 ry 0 rz -89.99 deg; joints [86.849, 39.666, -19.034, -0.718, -59.675, 93.452]
  MoveL 7 to (265.01, 36.7, 197.48) mm, rotated rx 168.69 ry 0 rz -89.99 deg; joints [86.872, 40.433, -18.579, -0.709, -60.131, 93.421]
  MoveL 8 to (252.92, 36.7, 196.02) mm, rotated rx 168.69 ry 0 rz -89.99 deg; joints [86.922, 42.216, -17.52, -0.691, -61.189, 93.352]
  MoveL 9 to (225.62, 36.7, 191.52) mm, rotated rx 168.69 ry 0 rz -89.99 deg; joints [87.028, 46.499, -14.955, -0.652, -63.753, 93.202]
  MoveL 10 to (214.97, 36.7, 189.31) mm, rotated rx 168.69 ry 0 rz -89.99 deg; joints [87.068, 48.285, -13.867, -0.637, -64.839, 93.146]
  MoveL 11 to (209.04, 36.7, 187.96) mm, rotated rx 168.69 ry 0 rz -89.99 deg; joints [87.09, 49.317, -13.233, -0.629, -65.473, 93.115]
  MoveL 12 to (205.72, 36.7, 187.17) mm, rotated rx 168.69 ry 0 rz -89.99 deg; joints [87.102, 49.905, -12.869, -0.625, -65.837, 93.098]
  MoveL 13 to (203.61, 36.7, 186.65) mm, rotated rx 168.69 ry 0 rz -89.99 deg; joints [87.109, 50.283, -12.634, -0.622, -66.072, 93.087]
  MoveL 14 to (201.54, 36.7, 186.06) mm, rotated rx 168.69 ry 0 rz -89.99 deg; joints [87.117, 50.662, -12.407, -0.619, -66.299, 93.076]
  MoveL 15 to (199.36, 36.7, 184) mm, rotated rx 168.69 ry 0 rz -89.99 deg; joints [87.124, 51.096, -12.336, -0.617, -66.37, 93.067]
  MoveL 16 to (198.9, 36.7, 182.55) mm, rotated rx 168.69 ry 0 rz -89.99 deg; joints [87.126, 51.212, -12.44, -0.618, -66.266, 93.067]
  MoveL 17 to (198.86, 36.7, 181.03) mm, rotated rx 168.69 ry 0 rz -89.99 deg; joints [87.126, 51.256, -12.612, -0.618, -66.095, 93.069]
  MoveL 18 to (198.86, 36.7, 174.94) mm, rotated rx 168.69 ry 0 rz -89.99 deg; joints [87.126, 51.411, -13.32, -0.622, -65.387, 93.077]
  MoveL 19 to (198.86, 36.7, 162.78) mm, rotated rx 168.69 ry 0 rz -89.99 deg; joints [87.126, 51.756, -14.71, -0.629, -63.996, 93.094]
  Establecer velocidad (1000.0 mm/s)
  MoveL 20 to (198.86, 36.7, 162.78) mm, rotated rx 168.69 ry 0 rz -89.99 deg; joints [87.126, 51.756, -14.71, -0.629, -63.996, 93.094]
  MoveL 21 to (218.47, 36.7, 260.83) mm, rotated rx 168.69 ry 0 rz -89.99 deg; joints [87.055, 46.596, -5.404, -0.605, -73.302, 93.062]
  Establecer velocidad (1000.0 mm/s)
  MoveL 22 to (294.14, 36.7, 296.46) mm, rotated rx 168.69 ry 0 rz -89.99 deg; joints [86.744, 33.884, -9.121, -0.683, -69.59, 93.431]
  MoveL 23 to (274.53, 36.7, 198.4) mm, rotated rx 168.69 ry 0 rz -89.99 deg; joints [86.831, 39.07, -19.388, -0.724, -59.322, 93.477]
  MoveL 24 to (274.53, 36.7, 198.4) mm, rotated rx 168.69 ry 0 rz -89.99 deg; joints [86.831, 39.07, -19.388, -0.724, -59.322, 93.477]
  Establecer velocidad (50.0 mm/s)
  MoveL 25 to (290.09, 36.7, 200.41) mm, rotated rx 168.69 ry 0 rz -89.99 deg; joints [86.763, 36.878, -20.564, -0.749, -58.147, 93.57]
  MoveL 26 to (305.43, 36.7, 203.7) mm, rotated rx 168.69 ry 0 rz -89.99 deg; joints [86.693, 34.719, -21.471, -0.773, -57.241, 93.661]
  MoveL 27 to (320.47, 36.7, 208.25) mm, rotated rx 168.69 ry 0 rz -89.99 deg; joints [86.621, 32.587, -22.114, -0.796, -56.599, 93.752]
  MoveL 28 to (335.07, 36.7, 214.04) mm, rotated rx 168.69 ry 0 rz -89.99 deg; joints [86.548, 30.488, -22.491, -0.816, -56.223, 93.839]
  MoveL 29 to (352.88, 36.7, 223.12) mm, rotated rx 168.69 ry 0 rz -89.99 deg; joints [86.455, 27.871, -22.593, -0.839, -56.122, 93.944]
  MoveL 30 to (369.63, 36.7, 234.02) mm, rotated rx 168.69 ry 0 rz -89.99 deg; joints [86.362, 25.334, -22.282, -0.858, -56.434, 94.042]
  MoveL 31 to (385.16, 36.7, 246.62) mm, rotated rx 168.69 ry 0 rz -89.99 deg; joints [86.272, 22.905, -21.574, -0.872, -57.143, 94.129]
  MoveL 32 to (399.27, 36.7, 260.77) mm, rotated rx 168.69 ry 0 rz -89.99 deg; joints [86.186, 20.617, -20.492, -0.881, -58.226, 94.204]
  Establecer velocidad (1000.0 mm/s)
  MoveL 33 to (399.27, 36.7, 260.77) mm, rotated rx 168.69 ry 0 rz -89.99 deg; joints [86.186, 20.617, -20.492, -0.881, -58.226, 94.204]
  MoveL 34 to (418.88, 36.7, 358.83) mm, rotated rx 168.69 ry 0 rz -89.99 deg; joints [86.059, 15.893, -8.512, -0.823, -70.207, 94.143]
  Establecer velocidad (1000.0 mm/s)
  MoveL 35 to (520.11, 36.7, 358.83) mm, rotated rx 168.69 ry 0 rz -89.99 deg; joints [85.248, 2.727, -10.739, -1.006, -67.994, 95.037]
  MoveL 36 to (500.5, 36.7, 260.77) mm, rotated rx 168.69 ry 0 rz -89.99 deg; joints [85.431, 8.03, -23.893, -1.097, -54.838, 95.112]
  MoveL 37 to (500.5, 36.7, 260.77) mm, rotated rx 168.69 ry 0 rz -89.99 deg; joints [85.431, 8.03, -23.893, -1.097, -54.838, 95.112]
  Establecer velocidad (50.0 mm/s)
  MoveL 38 to (502.78, 36.7, 247.62) mm, rotated rx 168.69 ry 0 rz -89.99 deg; joints [85.411, 8.346, -25.747, -1.128, -52.985, 95.18]
  MoveL 39 to (505.34, 36.7, 234.52) mm, rotated rx 168.69 ry 0 rz -89.99 deg; joints [85.388, 8.683, -27.61, -1.163, -51.123, 95.253]
  MoveL 40 to (508.02, 36.7, 221.45) mm, rotated rx 168.69 ry 0 rz -89.99 deg; joints [85.363, 9.065, -29.486, -1.202, -49.248, 95.332]
  MoveL 41 to (509.41, 36.7, 208.78) mm, rotated rx 168.69 ry 0 rz -89.99 deg; joints [85.351, 9.638, -31.287, -1.239, -47.447, 95.398]
  MoveL 42 to (509.37, 36.7, 196.07) mm, rotated rx 168.69 ry 0 rz -89.99 deg; joints [85.351, 10.442, -33.07, -1.276, -45.665, 95.451]
  MoveL 43 to (507.91, 36.7, 183.53) mm, rotated rx 168.69 ry 0 rz -89.99 deg; joints [85.365, 11.454, -34.793, -1.311, -43.942, 95.49]
  MoveL 44 to (505.04, 36.7, 171.19) mm, rotated rx 168.69 ry 0 rz -89.99 deg; joints [85.391, 12.662, -36.439, -1.345, -42.295, 95.515]
  Establecer velocidad (1000.0 mm/s)
  MoveL 45 to (505.04, 36.7, 171.19) mm, rotated rx 168.69 ry 0 rz -89.99 deg; joints [85.391, 12.662, -36.439, -1.345, -42.295, 95.515]
  MoveL 46 to (524.65, 36.7, 269.25) mm, rotated rx 168.69 ry 0 rz -89.99 deg; joints [85.205, 4.628, -23.09, -1.14, -55.645, 95.346]

--- program final (robot Fanuc LR Mate 200iD/7L) ---
  Llamar home
  Llamar reset
  Llamar c1 recoger
  Llamar poscharolamesa
  Llamar home
  Llamar iman izquierdo
  Llamar iman derecho
  Llamar recoger cepillo limpi...: recoger cepillo limpieza
  Llamar platizq
  Llamar parrizq
  Llamar platder
  Llamar parrder
  Llamar dejar cepillo limpieza
  Llamar recoger cera
  Llamar cerlatizq
  Llamar carribizq
  Llamar cerlatder
  Llamar cerarribder
  Llamar talonder
  Llamar dejar  cera
  Llamar recoger cepillo cera
  Llamar parrizq
  Llamar platder
  Llamar parrder
  Llamar dejar cepillo cera
  Llamar dejar iman izquierdo
  Llamar home
  Llamar dejar iman derecho
  Llamar pick charola
  Llamar c1 entregar

--- program cerlatizq (robot Fanuc LR Mate 200iD/7L) ---
  Suave(1)
  Establecer velocidad (1000.0 mm/s)
  Est. Ref.: RobotiQ 2F-140 Gripper (Mechanism) Base
  Est. herr: Tool 1
  Mostrar Tool 1
  MoveJ 1 to (287.12, 75.14, 245.65) mm, rotated rx 163.98 ry -47.25 rz -95.6 deg; joints [66.099, 43.658, -21.947, -52.065, -73.655, 119.467]
  MoveL 2 to (287.12, 75.14, 245.65) mm, rotated rx 163.98 ry -47.25 rz -95.6 deg; joints [66.099, 43.658, -21.947, -52.065, -73.655, 119.467]
  MoveL 3 to (267.51, 75.14, 147.59) mm, rotated rx 163.98 ry -47.25 rz -95.6 deg; joints [66.687, 51.246, -29.998, -54.435, -68.408, 125.951]
  MoveL 4 to (267.51, 75.14, 147.59) mm, rotated rx 163.98 ry -47.25 rz -95.6 deg; joints [66.687, 51.246, -29.998, -54.435, -68.408, 125.951]
  Establecer velocidad (50.0 mm/s)
  MoveL 5 to (279.24, 76.13, 147.59) mm, rotated rx 163.98 ry -47.25 rz -95.6 deg; joints [66.271, 49.909, -31.196, -54.697, -68.005, 127.226]
  MoveL 6 to (291.05, 76.12, 147.59) mm, rotated rx 163.98 ry -47.25 rz -95.6 deg; joints [65.911, 48.556, -32.397, -54.98, -67.564, 128.477]
  MoveL 7 to (302.8, 75.1, 147.59) mm, rotated rx 163.98 ry -47.25 rz -95.6 deg; joints [65.612, 47.199, -33.589, -55.286, -67.088, 129.692]
  MoveL 8 to (314.39, 73.1, 147.59) mm, rotated rx 163.98 ry -47.25 rz -95.6 deg; joints [65.38, 45.849, -34.764, -55.616, -66.58, 130.863]
  MoveL 9 to (325.74, 70.14, 148.13) mm, rotated rx 163.98 ry -47.25 rz -95.6 deg; joints [65.218, 44.473, -35.86, -55.952, -66.073, 131.934]
  MoveL 10 to (337.45, 66.21, 149.8) mm, rotated rx 163.98 ry -47.25 rz -95.6 deg; joints [65.11, 42.964, -36.872, -56.287, -65.581, 132.908]
  MoveL 11 to (349.04, 62.74, 152.6) mm, rotated rx 163.98 ry -47.25 rz -95.6 deg; joints [64.967, 41.432, -37.696, -56.544, -65.22, 133.732]
  MoveL 12 to (360.53, 59.92, 156.52) mm, rotated rx 163.98 ry -47.25 rz -95.6 deg; joints [64.774, 39.875, -38.324, -56.707, -65.001, 134.403]
  MoveL 13 to (372.2, 57.65, 160.01) mm, rotated rx 163.98 ry -47.25 rz -95.6 deg; joints [64.525, 38.371, -38.946, -56.845, -64.823, 135.095]
  MoveL 14 to (384.15, 55.93, 162.34) mm, rotated rx 163.98 ry -47.25 rz -95.6 deg; joints [64.214, 36.961, -39.653, -56.99, -64.639, 135.895]
  MoveL 15 to (396.39, 54.8, 163.5) mm, rotated rx 163.98 ry -47.25 rz -95.6 deg; joints [63.833, 35.651, -40.452, -57.139, -64.449, 136.813]
  MoveL 16 to (409.71, 54.28, 163.62) mm, rotated rx 163.98 ry -47.25 rz -95.6 deg; joints [63.347, 34.363, -41.387, -57.294, -64.252, 137.905]
  MoveL 17 to (423.03, 54.49, 163.62) mm, rotated rx 163.98 ry -47.25 rz -95.6 deg; joints [62.782, 33.136, -42.278, -57.39, -64.125, 138.992]
  MoveL 18 to (436.36, 54.49, 163.62) mm, rotated rx 163.98 ry -47.25 rz -95.6 deg; joints [62.213, 31.916, -43.147, -57.469, -64.01, 140.056]
  MoveL 19 to (449.69, 54.49, 163.62) mm, rotated rx 163.98 ry -47.25 rz -95.6 deg; joints [61.621, 30.712, -43.985, -57.519, -63.922, 141.099]
  MoveL 20 to (463.02, 54.49, 163.62) mm, rotated rx 163.98 ry -47.25 rz -95.6 deg; joints [61.005, 29.523, -44.794, -57.538, -63.859, 142.122]
  MoveL 21 to (471.35, 54.49, 163.62) mm, rotated rx 163.98 ry -47.25 rz -95.6 deg; joints [60.608, 28.786, -45.284, -57.535, -63.832, 142.751]
  MoveL 22 to (479.68, 54.49, 163.62) mm, rotated rx 163.98 ry -47.25 rz -95.6 deg; joints [60.201, 28.055, -45.764, -57.518, -63.815, 143.373]
  MoveL 23 to (488.01, 54.49, 163.62) mm, rotated rx 163.98 ry -47.25 rz -95.6 deg; joints [59.783, 27.328, -46.233, -57.489, -63.808, 143.987]
  MoveL 24 to (496.42, 54.24, 163.62) mm, rotated rx 163.98 ry -47.25 rz -95.6 deg; joints [59.372, 26.587, -46.703, -57.461, -63.794, 144.598]
  MoveL 25 to (502.24, 52.81, 163.62) mm, rotated rx 163.98 ry -47.25 rz -95.6 deg; joints [59.194, 26.011, -47.062, -57.512, -63.704, 145.01]
  MoveL 26 to (507.87, 49.97, 163.62) mm, rotated rx 163.98 ry -47.25 rz -95.6 deg; joints [59.147, 25.381, -47.449, -57.648, -63.523, 145.393]
  MoveL 27 to (512.8, 45.83, 163.62) mm, rotated rx 163.98 ry -47.25 rz -95.6 deg; joints [59.255, 24.744, -47.833, -57.872, -63.256, 145.713]
  MoveL 28 to (516.61, 40.68, 163.62) mm, rotated rx 163.98 ry -47.25 rz -95.6 deg; joints [59.52, 24.152, -48.184, -58.172, -62.92, 145.942]
  MoveL 29 to (519.08, 34.98, 163.62) mm, rotated rx 163.98 ry -47.25 rz -95.6 deg; joints [59.915, 23.65, -48.477, -58.525, -62.543, 146.067]
  MoveL 30 to (520.17, 29.21, 163.62) mm, rotated rx 163.98 ry -47.25 rz -95.6 deg; joints [60.399, 23.267, -48.698, -58.899, -62.155, 146.092]
  MoveL 31 to (520.26, 23.64, 163.62) mm, rotated rx 163.98 ry -47.25 rz -95.6 deg; joints [60.923, 22.986, -48.858, -59.272, -61.776, 146.047]
  MoveL 32 to (520.26, 18.08, 163.62) mm, rotated rx 163.98 ry -47.25 rz -95.6 deg; joints [61.456, 22.718, -49.01, -59.649, -61.398, 145.993]
  MoveL 33 to (519.72, 12.41, 163.62) mm, rotated rx 163.98 ry -47.25 rz -95.6 deg; joints [62.034, 22.496, -49.134, -60.04, -61.008, 145.898]
  MoveL 34 to (517.87, 6.62, 163.62) mm, rotated rx 163.98 ry -47.25 rz -95.6 deg; joints [62.696, 22.391, -49.192, -60.448, -60.603, 145.71]
  MoveL 35 to (514.63, 1.16, 163.62) mm, rotated rx 163.98 ry -47.25 rz -95.6 deg; joints [63.395, 22.433, -49.169, -60.839, -60.217, 145.429]
  MoveL 36 to (510.14, -3.47, 163.62) mm, rotated rx 163.98 ry -47.25 rz -95.6 deg; joints [64.071, 22.631, -49.058, -61.171, -59.883, 145.07]
  MoveL 37 to (504.76, -6.9, 163.62) mm, rotated rx 163.98 ry -47.25 rz -95.6 deg; joints [64.665, 22.969, -48.867, -61.412, -59.632, 144.66]
  MoveL 38 to (498.97, -8.95, 163.62) mm, rotated rx 163.98 ry -47.25 rz -95.6 deg; joints [65.134, 23.408, -48.616, -61.548, -59.481, 144.233]
  MoveL 39 to (491.37, -9.65, 163.62) mm, rotated rx 163.98 ry -47.25 rz -95.6 deg; joints [65.544, 24.07, -48.232, -61.579, -59.424, 143.689]
  MoveL 40 to (483.97, -9.65, 163.62) mm, rotated rx 163.98 ry -47.25 rz -95.6 deg; joints [65.868, 24.746, -47.831, -61.551, -59.425, 143.16]
  MoveL 41 to (476.56, -9.65, 163.62) mm, rotated rx 163.98 ry -47.25 rz -95.6 deg; joints [66.184, 25.425, -47.422, -61.512, -59.433, 142.624]
  MoveL 42 to (469.16, -9.65, 163.62) mm, rotated rx 163.98 ry -47.25 rz -95.6 deg; joints [66.492, 26.105, -47.003, -61.462, -59.448, 142.081]
  MoveL 43 to (461.75, -9.65, 163.62) mm, rotated rx 163.98 ry -47.25 rz -95.6 deg; joints [66.793, 26.788, -46.576, -61.401, -59.472, 141.531]
  MoveL 44 to (454.35, -9.65, 163.62) mm, rotated rx 163.98 ry -47.25 rz -95.6 deg; joints [67.087, 27.473, -46.14, -61.331, -59.503, 140.974]
  MoveL 45 to (439.69, -9.65, 163.62) mm, rotated rx 163.98 ry -47.25 rz -95.6 deg; joints [67.648, 28.838, -45.249, -61.163, -59.588, 139.85]
  MoveL 46 to (425.03, -9.65, 163.62) mm, rotated rx 163.98 ry -47.25 rz -95.6 deg; joints [68.183, 30.216, -44.324, -60.958, -59.703, 138.698]
  MoveL 47 to (410.37, -10.14, 163.62) mm, rotated rx 163.98 ry -47.25 rz -95.6 deg; joints [68.737, 31.59, -43.375, -60.745, -59.816, 137.513]
  MoveL 48 to (395.79, -11.63, 163.47) mm, rotated rx 163.98 ry -47.25 rz -95.6 deg; joints [69.351, 32.95, -42.438, -60.56, -59.884, 136.314]
  MoveL 49 to (383.65, -13.65, 162.27) mm, rotated rx 163.98 ry -47.25 rz -95.6 deg; joints [69.909, 34.153, -41.77, -60.479, -59.852, 135.407]
  MoveL 50 to (371.81, -16.31, 159.91) mm, rotated rx 163.98 ry -47.25 rz -95.6 deg; joints [70.493, 35.406, -41.239, -60.471, -59.733, 134.622]
  MoveL 51 to (360.26, -19.45, 156.42) mm, rotated rx 163.98 ry -47.25 rz -95.6 deg; joints [71.09, 36.711, -40.832, -60.526, -59.541, 133.955]
  MoveL 52 to (348.77, -22.13, 152.52) mm, rotated rx 163.98 ry -47.25 rz -95.6 deg; joints [71.631, 38.069, -40.426, -60.55, -59.384, 133.31]
  MoveL 53 to (336.98, -24.24, 149.71) mm, rotated rx 163.98 ry -47.25 rz -95.6 deg; joints [72.116, 39.403, -39.825, -60.445, -59.357, 132.489]
  MoveL 54 to (324.89, -25.75, 148.06) mm, rotated rx 163.98 ry -47.25 rz -95.6 deg; joints [72.546, 40.716, -39.025, -60.211, -59.464, 131.492]
  MoveL 55 to (313.84, -26.56, 147.59) mm, rotated rx 163.98 ry -47.25 rz -95.6 deg; joints [72.883, 41.875, -38.141, -59.893, -59.678, 130.45]
  MoveL 56 to (302.71, -26.83, 147.59) mm, rotated rx 163.98 ry -47.25 rz -95.6 deg; joints [73.17, 43.047, -37.157, -59.508, -59.978, 129.335]
  MoveL 57 to (291.57, -26.83, 147.59) mm, rotated rx 163.98 ry -47.25 rz -95.6 deg; joints [73.427, 44.252, -36.135, -59.097, -60.322, 128.2]
  MoveL 58 to (280.45, -26.23, 147.59) mm, rotated rx 163.98 ry -47.25 rz -95.6 deg; joints [73.632, 45.501, -35.063, -58.649, -60.734, 127.048]
  MoveL 59 to (269.47, -24.36, 147.59) mm, rotated rx 163.98 ry -47.25 rz -95.6 deg; joints [73.732, 46.805, -33.932, -58.147, -61.256, 125.897]
  MoveL 60 to (258.79, -21.23, 147.79) mm, rotated rx 163.98 ry -47.25 rz -95.6 deg; joints [73.731, 48.137, -32.734, -57.598, -61.894, 124.743]
  MoveL 61 to (248.6, -16.93, 148.47) mm, rotated rx 163.98 ry -47.25 rz -95.6 deg; joints [73.635, 49.46, -31.461, -57.007, -62.65, 123.583]
  MoveL 62 to (238.92, -11.46, 149.55) mm, rotated rx 163.98 ry -47.25 rz -95.6 deg; joints [73.448, 50.78, -30.121, -56.387, -63.52, 122.426]
  MoveL 63 to (230.02, -4.98, 150.92) mm, rotated rx 163.98 ry -47.25 rz -95.6 deg; joints [73.178, 52.074, -28.753, -55.765, -64.478, 121.309]
  MoveL 64 to (225.07, -0.64, 151.85) mm, rotated rx 163.98 ry -47.25 rz -95.6 deg; joints [72.98, 52.835, -27.928, -55.397, -65.089, 120.665]
  MoveL 65 to (220.43, 4.03, 152.83) mm, rotated rx 163.98 ry -47.25 rz -95.6 deg; joints [72.756, 53.588, -27.101, -55.034, -65.724, 120.043]
  MoveL 66 to (216.12, 9.07, 153.83) mm, rotated rx 163.98 ry -47.25 rz -95.6 deg; joints [72.502, 54.331, -26.278, -54.68, -66.383, 119.45]
  MoveL 67 to (212.91, 14.88, 154.63) mm, rotated rx 163.98 ry -47.25 rz -95.6 deg; joints [72.177, 54.988, -25.562, -54.359, -67.037, 119]
  MoveL 68 to (211.24, 21.32, 155.07) mm, rotated rx 163.98 ry -47.25 rz -95.6 deg; joints [71.778, 55.495, -25.034, -54.098, -67.638, 118.764]
  MoveL 69 to (211.02, 28.77, 155.13) mm, rotated rx 163.98 ry -47.25 rz -95.6 deg; joints [71.283, 55.877, -24.674, -53.879, -68.213, 118.735]
  MoveL 70 to (211.6, 36.19, 154.97) mm, rotated rx 163.98 ry -47.25 rz -95.6 deg; joints [70.774, 56.169, -24.429, -53.697, -68.732, 118.816]
  MoveL 71 to (213.49, 43.36, 154.48) mm, rotated rx 163.98 ry -47.25 rz -95.6 deg; joints [70.253, 56.288, -24.389, -53.578, -69.137, 119.083]
  MoveL 72 to (216.59, 50.02, 153.71) mm, rotated rx 163.98 ry -47.25 rz -95.6 deg; joints [69.737, 56.233, -24.552, -53.519, -69.418, 119.522]
  MoveL 73 to (220.83, 56.02, 152.74) mm, rotated rx 163.98 ry -47.25 rz -95.6 deg; joints [69.235, 56.004, -24.904, -53.517, -69.575, 120.114]
  MoveL 74 to (226.05, 61.17, 151.66) mm, rotated rx 163.98 ry -47.25 rz -95.6 deg; joints [68.763, 55.611, -25.423, -53.565, -69.611, 120.83]
  MoveL 75 to (232.09, 65.31, 150.57) mm, rotated rx 163.98 ry -47.25 rz -95.6 deg; joints [68.331, 55.067, -26.081, -53.661, -69.533, 121.642]
  MoveL 76 to (238.78, 68.33, 149.57) mm, rotated rx 163.98 ry -47.25 rz -95.6 deg; joints [67.953, 54.391, -26.849, -53.8, -69.352, 122.516]
  MoveL 77 to (245.8, 70.6, 148.73) mm, rotated rx 163.98 ry -47.25 rz -95.6 deg; joints [67.61, 53.642, -27.655, -53.958, -69.123, 123.405]
  MoveL 78 to (252.94, 72.49, 148.12) mm, rotated rx 163.98 ry -47.25 rz -95.6 deg; joints [67.284, 52.87, -28.45, -54.116, -68.889, 124.274]
  MoveL 79 to (260.17, 74.01, 147.74) mm, rotated rx 163.98 ry -47.25 rz -95.6 deg; joints [66.977, 52.071, -29.231, -54.275, -68.65, 125.123]
  MoveL 80 to (267.51, 75.14, 147.59) mm, rotated rx 163.98 ry -47.25 rz -95.6 deg; joints [66.687, 51.246, -29.998, -54.435, -68.408, 125.951]
  Establecer velocidad (1000.0 mm/s)
  MoveL 81 to (267.51, 75.14, 147.59) mm, rotated rx 163.98 ry -47.25 rz -95.6 deg; joints [66.687, 51.246, -29.998, -54.435, -68.408, 125.951]
  MoveL 82 to (287.12, 75.14, 245.65) mm, rotated rx 163.98 ry -47.25 rz -95.6 deg; joints [66.099, 43.658, -21.947, -52.065, -73.655, 119.467]
  Establecer velocidad (1000.0 mm/s)
  MoveL 83 to (478.44, -9.84, 310.93) mm, rotated rx 163.98 ry -47.25 rz -95.6 deg; joints [66.122, 14.485, -28.093, -53.684, -69.926, 124.612]
  MoveL 84 to (458.83, -9.84, 212.87) mm, rotated rx 163.98 ry -47.25 rz -95.6 deg; joints [66.927, 22.941, -40.165, -58.393, -62.607, 135.136]
  MoveL 85 to (458.83, -9.84, 212.87) mm, rotated rx 163.98 ry -47.25 rz -95.6 deg; joints [66.927, 22.941, -40.165, -58.393, -62.607, 135.136]
  Establecer velocidad (50.0 mm/s)
  MoveL 86 to (478.99, -8.87, 212.87) mm, rotated rx 163.98 ry -47.25 rz -95.6 deg; joints [66.006, 20.974, -41.113, -58.401, -62.705, 136.457]
  MoveL 87 to (499, -6.07, 212.87) mm, rotated rx 163.98 ry -47.25 rz -95.6 deg; joints [64.85, 19.119, -41.941, -58.229, -63.006, 137.761]
  MoveL 88 to (505.5, -4.27, 212.87) mm, rotated rx 163.98 ry -47.25 rz -95.6 deg; joints [64.371, 18.562, -42.177, -58.105, -63.184, 138.196]
  MoveL 89 to (511.4, -1.08, 212.87) mm, rotated rx 163.98 ry -47.25 rz -95.6 deg; joints [63.774, 18.134, -42.355, -57.896, -63.465, 138.626]
  MoveL 90 to (516.51, 3.32, 212.87) mm, rotated rx 163.98 ry -47.25 rz -95.6 deg; joints [63.088, 17.848, -42.471, -57.616, -63.831, 139.037]
  MoveL 91 to (520.5, 8.74, 212.87) mm, rotated rx 163.98 ry -47.25 rz -95.6 deg; joints [62.352, 17.732, -42.518, -57.28, -64.263, 139.406]
  MoveL 92 to (522.96, 15, 212.87) mm, rotated rx 163.98 ry -47.25 rz -95.6 deg; joints [61.613, 17.816, -42.484, -56.909, -64.739, 139.703]
  MoveL 93 to (523.6, 21.65, 212.87) mm, rotated rx 163.98 ry -47.25 rz -95.6 deg; joints [60.935, 18.105, -42.367, -56.534, -65.222, 139.897]
  MoveL 94 to (523.41, 27, 212.87) mm, rotated rx 163.98 ry -47.25 rz -95.6 deg; joints [60.434, 18.409, -42.241, -56.242, -65.6, 140.008]
  MoveL 95 to (522.19, 32.14, 212.87) mm, rotated rx 163.98 ry -47.25 rz -95.6 deg; joints [60.013, 18.804, -42.076, -55.977, -65.951, 140.048]
  MoveL 96 to (519.93, 36.95, 212.87) mm, rotated rx 163.98 ry -47.25 rz -95.6 deg; joints [59.685, 19.281, -41.872, -55.743, -66.268, 140.014]
  MoveL 97 to (516.79, 41.19, 212.87) mm, rotated rx 163.98 ry -47.25 rz -95.6 deg; joints [59.463, 19.81, -41.641, -55.552, -66.535, 139.907]
  MoveL 98 to (512.95, 44.85, 212.87) mm, rotated rx 163.98 ry -47.25 rz -95.6 deg; joints [59.336, 20.373, -41.389, -55.402, -66.756, 139.74]
  MoveL 99 to (507.06, 48.58, 212.87) mm, rotated rx 163.98 ry -47.25 rz -95.6 deg; joints [59.315, 21.131, -41.04, -55.269, -66.967, 139.438]
  MoveL 100 to (500.41, 50.78, 212.87) mm, rotated rx 163.98 ry -47.25 rz -95.6 deg; joints [59.47, 21.875, -40.688, -55.22, -67.072, 139.051]
  MoveL 101 to (493.51, 51.93, 212.87) mm, rotated rx 163.98 ry -47.25 rz -95.6 deg; joints [59.726, 22.585, -40.342, -55.219, -67.109, 138.622]
  MoveL 102 to (486.58, 52.86, 212.87) mm, rotated rx 163.98 ry -47.25 rz -95.6 deg; joints [59.997, 23.288, -39.992, -55.223, -67.139, 138.181]
  MoveL 103 to (479.62, 53.58, 212.87) mm, rotated rx 163.98 ry -47.25 rz -95.6 deg; joints [60.281, 23.983, -39.636, -55.229, -67.162, 137.729]
  MoveL 104 to (472.64, 54.1, 212.87) mm, rotated rx 163.98 ry -47.25 rz -95.6 deg; joints [60.578, 24.672, -39.276, -55.238, -67.179, 137.266]
  MoveL 105 to (456.16, 54.53, 212.87) mm, rotated rx 163.98 ry -47.25 rz -95.6 deg; joints [61.321, 26.267, -38.411, -55.267, -67.196, 136.138]
  MoveL 106 to (439.68, 53.94, 212.87) mm, rotated rx 163.98 ry -47.25 rz -95.6 deg; joints [62.113, 27.827, -37.526, -55.298, -67.188, 134.963]
  MoveL 107 to (429.96, 52.89, 212.87) mm, rotated rx 163.98 ry -47.25 rz -95.6 deg; joints [62.62, 28.722, -37.002, -55.327, -67.154, 134.246]
  MoveL 108 to (420.38, 51.24, 212.87) mm, rotated rx 163.98 ry -47.25 rz -95.6 deg; joints [63.157, 29.581, -36.486, -55.366, -67.093, 133.52]
  MoveL 109 to (410.84, 49.74, 212.87) mm, rotated rx 163.98 ry -47.25 rz -95.6 deg; joints [63.668, 30.455, -35.952, -55.383, -67.058, 132.788]
  MoveL 110 to (401.14, 49.84, 212.87) mm, rotated rx 163.98 ry -47.25 rz -95.6 deg; joints [64.043, 31.433, -35.34, -55.316, -67.155, 132.053]
  MoveL 111 to (391.44, 49.99, 212.87) mm, rotated rx 163.98 ry -47.25 rz -95.6 deg; joints [64.405, 32.423, -34.707, -55.234, -67.272, 131.306]
  MoveL 112 to (381.75, 49.97, 212.87) mm, rotated rx 163.98 ry -47.25 rz -95.6 deg; joints [64.77, 33.415, -34.059, -55.146, -67.394, 130.543]
  MoveL 113 to (377.34, 49.84, 212.87) mm, rotated rx 163.98 ry -47.25 rz -95.6 deg; joints [64.943, 33.864, -33.762, -55.107, -67.447, 130.191]
  MoveL 114 to (372.94, 49.58, 212.87) mm, rotated rx 163.98 ry -47.25 rz -95.6 deg; joints [65.123, 34.308, -33.465, -55.07, -67.494, 129.835]
  MoveL 115 to (368.55, 49.14, 212.87) mm, rotated rx 163.98 ry -47.25 rz -95.6 deg; joints [65.314, 34.745, -33.171, -55.038, -67.531, 129.474]
  MoveL 116 to (364.28, 48.09, 212.87) mm, rotated rx 163.98 ry -47.25 rz -95.6 deg; joints [65.546, 35.144, -32.9, -55.026, -67.527, 129.113]
  MoveL 117 to (360.68, 45.54, 212.87) mm, rotated rx 163.98 ry -47.25 rz -95.6 deg; joints [65.869, 35.402, -32.724, -55.077, -67.406, 128.789]
  MoveL 118 to (358.47, 42.59, 212.87) mm, rotated rx 163.98 ry -47.25 rz -95.6 deg; joints [66.173, 35.497, -32.659, -55.157, -67.233, 128.572]
  MoveL 119 to (357.27, 39.11, 212.87) mm, rotated rx 163.98 ry -47.25 rz -95.6 deg; joints [66.483, 35.463, -32.682, -55.27, -67.005, 128.431]
  MoveL 120 to (357.35, 35.44, 212.87) mm, rotated rx 163.98 ry -47.25 rz -95.6 deg; joints [66.765, 35.286, -32.803, -55.408, -66.741, 128.393]
  MoveL 121 to (359.01, 30.17, 212.87) mm, rotated rx 163.98 ry -47.25 rz -95.6 deg; joints [67.123, 34.871, -33.086, -55.629, -66.334, 128.462]
  MoveL 122 to (360.81, 24.94, 212.87) mm, rotated rx 163.98 ry -47.25 rz -95.6 deg; joints [67.475, 34.447, -33.372, -55.854, -65.929, 128.539]
  MoveL 123 to (360.26, 22.59, 212.87) mm, rotated rx 163.98 ry -47.25 rz -95.6 deg; joints [67.679, 34.403, -33.401, -55.934, -65.771, 128.461]
  MoveL 124 to (359.56, 20.23, 212.87) mm, rotated rx 163.98 ry -47.25 rz -95.6 deg; joints [67.889, 34.374, -33.421, -56.013, -65.616, 128.371]
  MoveL 125 to (358.88, 17.87, 212.87) mm, rotated rx 163.98 ry -47.25 rz -95.6 deg; joints [68.098, 34.345, -33.44, -56.091, -65.46, 128.282]
  MoveL 126 to (358.22, 15.51, 212.87) mm, rotated rx 163.98 ry -47.25 rz -95.6 deg; joints [68.308, 34.316, -33.46, -56.17, -65.303, 128.192]
  MoveL 127 to (357.56, 13.14, 212.87) mm, rotated rx 163.98 ry -47.25 rz -95.6 deg; joints [68.518, 34.285, -33.481, -56.248, -65.147, 128.104]
  MoveL 128 to (357.19, 10.73, 212.87) mm, rotated rx 163.98 ry -47.25 rz -95.6 deg; joints [68.722, 34.224, -33.521, -56.333, -64.982, 128.037]
  MoveL 129 to (357.76, 5.92, 212.87) mm, rotated rx 163.98 ry -47.25 rz -95.6 deg; joints [69.091, 33.965, -33.694, -56.525, -64.631, 128.009]
  MoveL 130 to (359.87, 1.54, 212.87) mm, rotated rx 163.98 ry -47.25 rz -95.6 deg; joints [69.38, 33.562, -33.962, -56.729, -64.283, 128.11]
  MoveL 131 to (363.08, -2.1, 212.87) mm, rotated rx 163.98 ry -47.25 rz -95.6 deg; joints [69.579, 33.076, -34.282, -56.927, -63.97, 128.307]
  MoveL 132 to (367.29, -4.48, 212.87) mm, rotated rx 163.98 ry -47.25 rz -95.6 deg; joints [69.646, 32.534, -34.634, -57.095, -63.732, 128.604]
  MoveL 133 to (372.09, -5.28, 212.87) mm, rotated rx 163.98 ry -47.25 rz -95.6 deg; joints [69.564, 31.996, -34.981, -57.211, -63.6, 128.969]
  MoveL 134 to (376.94, -5.73, 212.87) mm, rotated rx 163.98 ry -47.25 rz -95.6 deg; joints [69.451, 31.468, -35.317, -57.311, -63.496, 129.341]
  MoveL 135 to (381.8, -5.94, 212.87) mm, rotated rx 163.98 ry -47.25 rz -95.6 deg; joints [69.315, 30.95, -35.643, -57.399, -63.413, 129.714]
  MoveL 136 to (386.67, -5.99, 212.87) mm, rotated rx 163.98 ry -47.25 rz -95.6 deg; joints [69.164, 30.44, -35.96, -57.478, -63.346, 130.087]
  MoveL 137 to (391.54, -5.93, 212.87) mm, rotated rx 163.98 ry -47.25 rz -95.6 deg; joints [69.002, 29.936, -36.27, -57.549, -63.29, 130.458]
  MoveL 138 to (396.99, -5.79, 212.87) mm, rotated rx 163.98 ry -47.25 rz -95.6 deg; joints [68.81, 29.378, -36.609, -57.621, -63.239, 130.871]
  MoveL 139 to (402.44, -5.61, 212.87) mm, rotated rx 163.98 ry -47.25 rz -95.6 deg; joints [68.612, 28.824, -36.94, -57.687, -63.195, 131.28]
  MoveL 140 to (407.89, -5.44, 212.87) mm, rotated rx 163.98 ry -47.25 rz -95.6 deg; joints [68.412, 28.272, -37.266, -57.748, -63.156, 131.684]
  MoveL 141 to (413.34, -5.32, 212.87) mm, rotated rx 163.98 ry -47.25 rz -95.6 deg; joints [68.213, 27.719, -37.588, -57.808, -63.119, 132.084]
  MoveL 142 to (418.69, -6.35, 212.87) mm, rotated rx 163.98 ry -47.25 rz -95.6 deg; joints [68.115, 27.132, -37.925, -57.914, -63.005, 132.45]
  MoveL 143 to (424.09, -7.65, 212.87) mm, rotated rx 163.98 ry -47.25 rz -95.6 deg; joints [68.038, 26.53, -38.264, -58.03, -62.876, 132.809]
  MoveL 144 to (430.03, -8.99, 212.87) mm, rotated rx 163.98 ry -47.25 rz -95.6 deg; joints [67.944, 25.874, -38.628, -58.15, -62.747, 133.2]
  MoveL 145 to (434.74, -9.6, 212.87) mm, rotated rx 163.98 ry -47.25 rz -95.6 deg; joints [67.826, 25.372, -38.901, -58.221, -62.681, 133.515]
  MoveL 146 to (438.44, -9.81, 212.87) mm, rotated rx 163.98 ry -47.25 rz -95.6 deg; joints [67.708, 24.99, -39.106, -58.262, -62.651, 133.766]
  MoveL 147 to (441.88, -9.84, 212.87) mm, rotated rx 163.98 ry -47.25 rz -95.6 deg; joints [67.582, 24.642, -39.291, -58.29, -62.637, 134.001]
  MoveL 148 to (444.88, -9.84, 212.87) mm, rotated rx 163.98 ry -47.25 rz -95.6 deg; joints [67.469, 24.34, -39.45, -58.312, -62.628, 134.205]
  MoveL 149 to (448.72, -9.84, 212.87) mm, rotated rx 163.98 ry -47.25 rz -95.6 deg; joints [67.322, 23.954, -39.65, -58.337, -62.619, 134.464]
  MoveL 150 to (453.55, -9.84, 212.87) mm, rotated rx 163.98 ry -47.25 rz -95.6 deg; joints [67.135, 23.47, -39.898, -58.366, -62.611, 134.787]
  MoveL 151 to (458.83, -9.84, 212.87) mm, rotated rx 163.98 ry -47.25 rz -95.6 deg; joints [66.927, 22.941, -40.165, -58.393, -62.607, 135.136]
  Establecer velocidad (1000.0 mm/s)
  MoveL 152 to (458.83, -9.84, 212.87) mm, rotated rx 163.98 ry -47.25 rz -95.6 deg; joints [66.927, 22.941, -40.165, -58.393, -62.607, 135.136]
  MoveL 153 to (478.44, -9.84, 310.93) mm, rotated rx 163.98 ry -47.25 rz -95.6 deg; joints [66.122, 14.485, -28.093, -53.684, -69.926, 124.612]

--- program platder (robot Fanuc LR Mate 200iD/7L) ---
  Suave(1)
  Establecer velocidad (1000.0 mm/s)
  Est. Ref.: RobotiQ 2F-140 Gripper (Mechanism) Base
  Est. herr: Tool 1
  Mostrar Tool 1
  MoveJ 1 to (296.61, 215.99, 331.82) mm, rotated rx -178.1 ry -46.22 rz 172.02 deg; joints [70.53, 20.204, -21.641, -24.631, -25.021, 30.604]
  MoveL 2 to (296.61, 215.99, 331.82) mm, rotated rx -178.1 ry -46.22 rz 172.02 deg; joints [70.53, 20.204, -21.641, -24.631, -25.021, 30.604]
  MoveL 3 to (277, 215.99, 233.76) mm, rotated rx -178.1 ry -46.22 rz 172.02 deg; joints [71.13, 27.321, -32.848, -40.178, -15.178, 46.793]
  MoveL 4 to (277, 215.99, 233.76) mm, rotated rx -178.1 ry -46.22 rz 172.02 deg; joints [71.13, 27.321, -32.848, -40.178, -15.178, 46.793]
  Establecer velocidad (50.0 mm/s)
  MoveL 5 to (288.59, 217.34, 233.76) mm, rotated rx -178.1 ry -46.22 rz 172.02 deg; joints [70.66, 26.118, -33.49, -42.595, -14.956, 49.562]
  MoveL 6 to (300.24, 217.49, 233.76) mm, rotated rx -178.1 ry -46.22 rz 172.02 deg; joints [70.28, 24.87, -34.132, -44.92, -14.711, 52.186]
  MoveL 7 to (311.9, 217.39, 233.76) mm, rotated rx -178.1 ry -46.22 rz 172.02 deg; joints [69.908, 23.621, -34.748, -47.23, -14.505, 54.791]
  MoveL 8 to (323.52, 216.75, 233.96) mm, rotated rx -178.1 ry -46.22 rz 172.02 deg; joints [69.574, 22.346, -35.319, -49.404, -14.33, 57.234]
  MoveL 9 to (335.6, 215.45, 235.24) mm, rotated rx -178.1 ry -46.22 rz 172.02 deg; joints [69.272, 20.927, -35.752, -51.154, -14.241, 59.22]
  MoveL 10 to (347.37, 213.53, 237.67) mm, rotated rx -178.1 ry -46.22 rz 172.02 deg; joints [69.028, 19.433, -35.994, -52.242, -14.247, 60.491]
  MoveL 11 to (358.85, 211.05, 241.24) mm, rotated rx -178.1 ry -46.22 rz 172.02 deg; joints [68.84, 17.862, -36.04, -52.638, -14.339, 61.013]
  MoveL 12 to (370.22, 208, 245.03) mm, rotated rx -178.1 ry -46.22 rz 172.02 deg; joints [68.705, 16.254, -36.013, -52.733, -14.442, 61.193]
  MoveL 13 to (381.87, 205.17, 247.71) mm, rotated rx -178.1 ry -46.22 rz 172.02 deg; joints [68.53, 14.692, -36.096, -53.217, -14.505, 61.8]
  MoveL 14 to (393.81, 202.97, 249.25) mm, rotated rx -178.1 ry -46.22 rz 172.02 deg; joints [68.269, 13.195, -36.292, -54.153, -14.559, 62.926]
  MoveL 15 to (406.9, 201.36, 249.64) mm, rotated rx -178.1 ry -46.22 rz 172.02 deg; joints [67.882, 11.671, -36.632, -55.681, -14.618, 64.742]
  MoveL 16 to (420.09, 200.57, 249.64) mm, rotated rx -178.1 ry -46.22 rz 172.02 deg; joints [67.382, 10.192, -36.978, -57.323, -14.761, 66.749]
  MoveL 17 to (433.3, 200.48, 249.64) mm, rotated rx -178.1 ry -46.22 rz 172.02 deg; joints [66.776, 8.734, -37.274, -58.863, -15.015, 68.722]
  MoveL 18 to (446.51, 200.48, 249.64) mm, rotated rx -178.1 ry -46.22 rz 172.02 deg; joints [66.128, 7.273, -37.526, -60.234, -15.331, 70.55]
  MoveL 19 to (459.72, 200.48, 249.64) mm, rotated rx -178.1 ry -46.22 rz 172.02 deg; joints [65.444, 5.803, -37.734, -61.421, -15.703, 72.215]
  MoveL 20 to (492.75, 200.48, 249.64) mm, rotated rx -178.1 ry -46.22 rz 172.02 deg; joints [63.564, 2.077, -38.053, -63.58, -16.872, 75.667]
  MoveL 21 to (498.39, 200.04, 249.64) mm, rotated rx -178.1 ry -46.22 rz 172.02 deg; joints [63.272, 1.408, -38.078, -63.809, -17.067, 76.095]
  MoveL 22 to (504.16, 198.3, 249.64) mm, rotated rx -178.1 ry -46.22 rz 172.02 deg; joints [63.125, 0.645, -38.096, -63.933, -17.163, 76.32]
  MoveL 23 to (509.62, 195.19, 249.64) mm, rotated rx -178.1 ry -46.22 rz 172.02 deg; joints [63.169, -0.171, -38.1, -63.923, -17.13, 76.28]
  MoveL 24 to (514.28, 190.82, 249.64) mm, rotated rx -178.1 ry -46.22 rz 172.02 deg; joints [63.429, -0.975, -38.09, -63.759, -16.951, 75.942]
  MoveL 25 to (517.77, 185.55, 249.64) mm, rotated rx -178.1 ry -46.22 rz 172.02 deg; joints [63.894, -1.698, -38.068, -63.444, -16.633, 75.313]
  MoveL 26 to (519.9, 179.84, 249.64) mm, rotated rx -178.1 ry -46.22 rz 172.02 deg; joints [64.518, -2.284, -38.043, -63, -16.205, 74.449]
  MoveL 27 to (520.69, 174.16, 249.64) mm, rotated rx -178.1 ry -46.22 rz 172.02 deg; joints [65.237, -2.703, -38.02, -62.465, -15.713, 73.432]
  MoveL 28 to (520.7, 168.65, 249.64) mm, rotated rx -178.1 ry -46.22 rz 172.02 deg; joints [65.991, -3.012, -38.001, -61.865, -15.196, 72.327]
  MoveL 29 to (520.68, 163.15, 249.64) mm, rotated rx -178.1 ry -46.22 rz 172.02 deg; joints [66.756, -3.308, -37.98, -61.19, -14.676, 71.142]
  MoveL 30 to (519.86, 157.46, 249.64) mm, rotated rx -178.1 ry -46.22 rz 172.02 deg; joints [67.602, -3.504, -37.966, -60.393, -14.101, 69.781]
  MoveL 31 to (517.7, 151.76, 249.64) mm, rotated rx -178.1 ry -46.22 rz 172.02 deg; joints [68.532, -3.521, -37.964, -59.462, -13.467, 68.233]
  MoveL 32 to (514.17, 146.5, 249.64) mm, rotated rx -178.1 ry -46.22 rz 172.02 deg; joints [69.471, -3.329, -37.979, -58.457, -12.825, 66.608]
  MoveL 33 to (509.48, 142.17, 249.64) mm, rotated rx -178.1 ry -46.22 rz 172.02 deg; joints [70.332, -2.934, -38.006, -57.471, -12.236, 65.055]
  MoveL 34 to (504, 139.09, 249.64) mm, rotated rx -178.1 ry -46.22 rz 172.02 deg; joints [71.039, -2.376, -38.038, -56.607, -11.751, 63.727]
  MoveL 35 to (497.41, 137.26, 249.64) mm, rotated rx -178.1 ry -46.22 rz 172.02 deg; joints [71.608, -1.621, -38.071, -55.874, -11.36, 62.62]
  MoveL 36 to (491.03, 136.98, 249.64) mm, rotated rx -178.1 ry -46.22 rz 172.02 deg; joints [71.938, -0.833, -38.092, -55.427, -11.133, 61.958]
  MoveL 37 to (484.74, 136.98, 249.64) mm, rotated rx -178.1 ry -46.22 rz 172.02 deg; joints [72.216, -0.049, -38.099, -54.991, -10.949, 61.338]
  MoveL 38 to (478.45, 136.98, 249.64) mm, rotated rx -178.1 ry -46.22 rz 172.02 deg; joints [72.486, 0.728, -38.094, -54.494, -10.779, 60.663]
  MoveL 39 to (472.16, 136.98, 249.64) mm, rotated rx -178.1 ry -46.22 rz 172.02 deg; joints [72.748, 1.501, -38.075, -53.937, -10.623, 59.931]
  MoveL 40 to (465.86, 136.98, 249.64) mm, rotated rx -178.1 ry -46.22 rz 172.02 deg; joints [73.003, 2.267, -38.043, -53.32, -10.48, 59.144]
  MoveL 41 to (459.57, 136.98, 249.64) mm, rotated rx -178.1 ry -46.22 rz 172.02 deg; joints [73.25, 3.029, -37.999, -52.643, -10.351, 58.301]
  MoveL 42 to (445.04, 136.98, 249.64) mm, rotated rx -178.1 ry -46.22 rz 172.02 deg; joints [73.796, 4.771, -37.852, -50.859, -10.105, 56.148]
  MoveL 43 to (430.51, 136.98, 249.64) mm, rotated rx -178.1 ry -46.22 rz 172.02 deg; joints [74.308, 6.489, -37.642, -48.787, -9.931, 53.725]
  MoveL 44 to (415.98, 137.19, 249.64) mm, rotated rx -178.1 ry -46.22 rz 172.02 deg; joints [74.764, 8.195, -37.372, -46.52, -9.845, 51.142]
  MoveL 45 to (401.45, 136.87, 249.62) mm, rotated rx -178.1 ry -46.22 rz 172.02 deg; joints [75.255, 9.867, -37.05, -43.906, -9.794, 48.188]
  MoveL 46 to (389.24, 135.91, 248.8) mm, rotated rx -178.1 ry -46.22 rz 172.02 deg; joints [75.723, 11.301, -36.857, -41.824, -9.681, 45.79]
  MoveL 47 to (377.31, 134.37, 246.8) mm, rotated rx -178.1 ry -46.22 rz 172.02 deg; joints [76.226, 12.763, -36.802, -40.106, -9.459, 43.741]
  MoveL 48 to (365.67, 132.27, 243.66) mm, rotated rx -178.1 ry -46.22 rz 172.02 deg; joints [76.761, 14.253, -36.878, -38.7, -9.128, 41.991]
  MoveL 49 to (354.28, 129.63, 239.67) mm, rotated rx -178.1 ry -46.22 rz 172.02 deg; joints [77.326, 15.755, -37.038, -37.408, -8.724, 40.341]
  MoveL 50 to (342.81, 126.37, 236.59) mm, rotated rx -178.1 ry -46.22 rz 172.02 deg; joints [77.934, 17.18, -37.035, -35.169, -8.439, 37.706]
  MoveL 51 to (331.26, 122.49, 234.64) mm, rotated rx -178.1 ry -46.22 rz 172.02 deg; joints [78.584, 18.517, -36.843, -31.894, -8.312, 34]
  MoveL 52 to (318.55, 118.92, 233.78) mm, rotated rx -178.1 ry -46.22 rz 172.02 deg; joints [79.201, 19.912, -36.416, -27.903, -8.435, 29.594]
  MoveL 53 to (305.52, 116.58, 233.76) mm, rotated rx -178.1 ry -46.22 rz 172.02 deg; joints [79.676, 21.315, -35.815, -24.165, -8.807, 25.53]
  MoveL 54 to (292.27, 115.5, 233.76) mm, rotated rx -178.1 ry -46.22 rz 172.02 deg; joints [80.013, 22.771, -35.151, -21.171, -9.314, 22.301]
  MoveL 55 to (278.98, 115.71, 233.76) mm, rotated rx -178.1 ry -46.22 rz 172.02 deg; joints [80.214, 24.261, -34.435, -18.92, -9.931, 19.902]
  MoveL 56 to (265.83, 117.19, 233.83) mm, rotated rx -178.1 ry -46.22 rz 172.02 deg; joints [80.287, 25.761, -33.665, -17.327, -10.644, 18.241]
  MoveL 57 to (257.77, 118.75, 234.18) mm, rotated rx -178.1 ry -46.22 rz 172.02 deg; joints [80.271, 26.679, -33.129, -16.573, -11.16, 17.482]
  MoveL 58 to (249.83, 120.77, 234.81) mm, rotated rx -178.1 ry -46.22 rz 172.02 deg; joints [80.211, 27.578, -32.546, -15.973, -11.734, 16.903]
  MoveL 59 to (242.03, 123.27, 235.72) mm, rotated rx -178.1 ry -46.22 rz 172.02 deg; joints [80.108, 28.461, -31.919, -15.511, -12.361, 16.487]
  MoveL 60 to (234.65, 126.69, 236.84) mm, rotated rx -178.1 ry -46.22 rz 172.02 deg; joints [79.921, 29.309, -31.269, -15.329, -13.03, 16.4]
  MoveL 61 to (228.08, 131.5, 238.05) mm, rotated rx -178.1 ry -46.22 rz 172.02 deg; joints [79.604, 30.096, -30.632, -15.553, -13.717, 16.799]
  MoveL 62 to (222.62, 137.49, 239.22) mm, rotated rx -178.1 ry -46.22 rz 172.02 deg; joints [79.176, 30.793, -30.047, -16.121, -14.381, 17.607]
  MoveL 63 to (218.41, 144.51, 240.22) mm, rotated rx -178.1 ry -46.22 rz 172.02 deg; joints [78.647, 31.387, -29.543, -16.988, -14.994, 18.774]
  MoveL 64 to (215.69, 152.2, 240.92) mm, rotated rx -178.1 ry -46.22 rz 172.02 deg; joints [78.044, 31.852, -29.159, -18.106, -15.518, 20.24]
  MoveL 65 to (214.75, 157.63, 241.17) mm, rotated rx -178.1 ry -46.22 rz 172.02 deg; joints [77.605, 32.086, -28.98, -18.986, -15.81, 21.375]
  MoveL 66 to (214.52, 163.15, 241.23) mm, rotated rx -178.1 ry -46.22 rz 172.02 deg; joints [77.149, 32.254, -28.869, -19.956, -16.048, 22.613]
  MoveL 67 to (214.62, 168.67, 241.2) mm, rotated rx -178.1 ry -46.22 rz 172.02 deg; joints [76.687, 32.395, -28.787, -20.942, -16.266, 23.872]
  MoveL 68 to (215.64, 174.03, 240.93) mm, rotated rx -178.1 ry -46.22 rz 172.02 deg; joints [76.221, 32.441, -28.799, -22.03, -16.405, 25.239]
  MoveL 69 to (218.69, 180.65, 240.16) mm, rotated rx -178.1 ry -46.22 rz 172.02 deg; joints [75.609, 32.32, -28.988, -23.66, -16.438, 27.247]
  MoveL 70 to (223.25, 186.3, 239.08) mm, rotated rx -178.1 ry -46.22 rz 172.02 deg; joints [75.041, 32.021, -29.332, -25.401, -16.332, 29.351]
  MoveL 71 to (228.32, 191.45, 238.01) mm, rotated rx -178.1 ry -46.22 rz 172.02 deg; joints [74.498, 31.659, -29.712, -27.163, -16.2, 31.465]
  MoveL 72 to (236.59, 198.41, 236.52) mm, rotated rx -178.1 ry -46.22 rz 172.02 deg; joints [73.72, 31.025, -30.317, -29.825, -15.99, 34.64]
  MoveL 73 to (245.7, 204.45, 235.26) mm, rotated rx -178.1 ry -46.22 rz 172.02 deg; joints [72.985, 30.275, -30.951, -32.508, -15.774, 37.819]
  MoveL 74 to (255.44, 209.41, 234.33) mm, rotated rx -178.1 ry -46.22 rz 172.02 deg; joints [72.307, 29.416, -31.59, -35.14, -15.566, 40.918]
  MoveL 75 to (265.68, 213.23, 233.83) mm, rotated rx -178.1 ry -46.22 rz 172.02 deg; joints [71.697, 28.453, -32.213, -37.66, -15.372, 43.867]
  Establecer velocidad (1000.0 mm/s)
  MoveL 76 to (265.68, 213.23, 233.83) mm, rotated rx -178.1 ry -46.22 rz 172.02 deg; joints [71.697, 28.453, -32.213, -37.66, -15.372, 43.867]
  MoveL 77 to (285.29, 213.23, 331.89) mm, rotated rx -178.1 ry -46.22 rz 172.02 deg; joints [71.123, 21.427, -21.158, -23.352, -25.238, 28.952]
  Establecer velocidad (1000.0 mm/s)
  MoveL 78 to (479.49, 200.65, 396.6) mm, rotated rx -178.1 ry -46.22 rz 172.02 deg; joints [64.329, -4.285, -16.18, -27.823, -32.517, 36.529]
  MoveL 79 to (459.88, 200.65, 298.54) mm, rotated rx -178.1 ry -46.22 rz 172.02 deg; joints [65.416, 2.348, -30.399, -43.435, -20.253, 53.353]
  MoveL 80 to (459.88, 200.65, 298.54) mm, rotated rx -178.1 ry -46.22 rz 172.02 deg; joints [65.416, 2.348, -30.399, -43.435, -20.253, 53.353]
  Establecer velocidad (50.0 mm/s)
  MoveL 81 to (479.73, 199.7, 298.54) mm, rotated rx -178.1 ry -46.22 rz 172.02 deg; joints [64.43, -0.023, -30.455, -44.671, -20.805, 55.207]
  MoveL 82 to (499.42, 196.95, 298.54) mm, rotated rx -178.1 ry -46.22 rz 172.02 deg; joints [63.59, -2.513, -30.391, -45.455, -21.362, 56.502]
  MoveL 83 to (505.83, 195.22, 298.54) mm, rotated rx -178.1 ry -46.22 rz 172.02 deg; joints [63.406, -3.383, -30.339, -45.552, -21.512, 56.706]
  MoveL 84 to (511.67, 192.13, 298.54) mm, rotated rx -178.1 ry -46.22 rz 172.02 deg; joints [63.428, -4.273, -30.27, -45.405, -21.547, 56.536]
  MoveL 85 to (516.74, 187.86, 298.54) mm, rotated rx -178.1 ry -46.22 rz 172.02 deg; joints [63.656, -5.149, -30.187, -45.018, -21.466, 55.997]
  MoveL 86 to (520.73, 182.58, 298.54) mm, rotated rx -178.1 ry -46.22 rz 172.02 deg; joints [64.096, -5.96, -30.096, -44.384, -21.262, 55.079]
  MoveL 87 to (523.25, 176.47, 298.54) mm, rotated rx -178.1 ry -46.22 rz 172.02 deg; joints [64.758, -6.639, -30.01, -43.49, -20.927, 53.766]
  MoveL 88 to (523.99, 169.9, 298.54) mm, rotated rx -178.1 ry -46.22 rz 172.02 deg; joints [65.614, -7.116, -29.944, -42.362, -20.47, 52.102]
  MoveL 89 to (523.68, 163.32, 298.54) mm, rotated rx -178.1 ry -46.22 rz 172.02 deg; joints [66.551, -7.448, -29.896, -41.096, -19.965, 50.255]
  MoveL 90 to (521.79, 157.05, 298.54) mm, rotated rx -178.1 ry -46.22 rz 172.02 deg; joints [67.548, -7.547, -29.881, -39.727, -19.417, 48.273]
  MoveL 91 to (518.32, 151.45, 298.54) mm, rotated rx -178.1 ry -46.22 rz 172.02 deg; joints [68.541, -7.389, -29.904, -38.337, -18.856, 46.279]
  MoveL 92 to (513.71, 146.76, 298.54) mm, rotated rx -178.1 ry -46.22 rz 172.02 deg; joints [69.459, -7.023, -29.957, -37.019, -18.328, 44.405]
  MoveL 93 to (508.37, 143.24, 298.54) mm, rotated rx -178.1 ry -46.22 rz 172.02 deg; joints [70.236, -6.495, -30.029, -35.881, -17.87, 42.799]
  MoveL 94 to (502.4, 140.97, 298.54) mm, rotated rx -178.1 ry -46.22 rz 172.02 deg; joints [70.852, -5.822, -30.112, -34.98, -17.493, 41.53]
  MoveL 95 to (496.16, 139.84, 298.54) mm, rotated rx -178.1 ry -46.22 rz 172.02 deg; joints [71.308, -5.063, -30.195, -34.322, -17.201, 40.6]
  MoveL 96 to (489.87, 138.92, 298.54) mm, rotated rx -178.1 ry -46.22 rz 172.02 deg; joints [71.723, -4.291, -30.268, -33.695, -16.94, 39.725]
  MoveL 97 to (473.76, 137.39, 298.54) mm, rotated rx -178.1 ry -46.22 rz 172.02 deg; joints [72.627, -2.297, -30.401, -32.206, -16.404, 37.695]
  MoveL 98 to (457.58, 136.96, 298.54) mm, rotated rx -178.1 ry -46.22 rz 172.02 deg; joints [73.329, -0.277, -30.453, -30.882, -16.042, 35.945]
  MoveL 99 to (442.87, 137.39, 298.54) mm, rotated rx -178.1 ry -46.22 rz 172.02 deg; joints [73.822, 1.567, -30.429, -29.807, -15.849, 34.568]
  MoveL 100 to (428.32, 139.01, 298.54) mm, rotated rx -178.1 ry -46.22 rz 172.02 deg; joints [74.136, 3.41, -30.337, -28.973, -15.796, 33.536]
  MoveL 101 to (414.04, 141.71, 298.54) mm, rotated rx -178.1 ry -46.22 rz 172.02 deg; joints [74.294, 5.234, -30.178, -28.36, -15.87, 32.815]
  MoveL 102 to (399.51, 141.55, 298.54) mm, rotated rx -178.1 ry -46.22 rz 172.02 deg; joints [74.777, 6.976, -29.964, -26.952, -15.866, 31.1]
  MoveL 103 to (384.97, 141.47, 298.54) mm, rotated rx -178.1 ry -46.22 rz 172.02 deg; joints [75.224, 8.707, -29.692, -25.531, -15.938, 29.391]
  MoveL 104 to (380.65, 141.58, 298.54) mm, rotated rx -178.1 ry -46.22 rz 172.02 deg; joints [75.338, 9.224, -29.599, -25.135, -15.98, 28.921]
  MoveL 105 to (376.33, 141.79, 298.54) mm, rotated rx -178.1 ry -46.22 rz 172.02 deg; joints [75.438, 9.742, -29.501, -24.765, -16.032, 28.485]
  MoveL 106 to (372.02, 142.16, 298.54) mm, rotated rx -178.1 ry -46.22 rz 172.02 deg; joints [75.519, 10.264, -29.397, -24.431, -16.097, 28.096]
  MoveL 107 to (367.77, 142.86, 298.54) mm, rotated rx -178.1 ry -46.22 rz 172.02 deg; joints [75.562, 10.789, -29.287, -24.178, -16.182, 27.81]
  MoveL 108 to (363.99, 144.91, 298.54) mm, rotated rx -178.1 ry -46.22 rz 172.02 deg; joints [75.446, 11.296, -29.175, -24.28, -16.325, 27.976]
  MoveL 109 to (361.54, 147.54, 298.54) mm, rotated rx -178.1 ry -46.22 rz 172.02 deg; joints [75.235, 11.666, -29.091, -24.63, -16.478, 28.447]
  MoveL 110 to (359.93, 150.76, 298.54) mm, rotated rx -178.1 ry -46.22 rz 172.02 deg; joints [74.941, 11.956, -29.023, -25.175, -16.648, 29.165]
  MoveL 111 to (359.47, 154.31, 298.54) mm, rotated rx -178.1 ry -46.22 rz 172.02 deg; joints [74.581, 12.123, -28.983, -25.888, -16.82, 30.093]
  MoveL 112 to (360.22, 157.83, 298.54) mm, rotated rx -178.1 ry -46.22 rz 172.02 deg; joints [74.19, 12.15, -28.977, -26.699, -16.977, 31.138]
  MoveL 113 to (361.37, 161.27, 298.54) mm, rotated rx -178.1 ry -46.22 rz 172.02 deg; joints [73.796, 12.131, -28.981, -27.515, -17.13, 32.191]
  MoveL 114 to (362.55, 164.7, 298.54) mm, rotated rx -178.1 ry -46.22 rz 172.02 deg; joints [73.402, 12.111, -28.986, -28.314, -17.287, 33.227]
  MoveL 115 to (362.88, 167.44, 298.54) mm, rotated rx -178.1 ry -46.22 rz 172.02 deg; joints [73.106, 12.169, -28.972, -28.877, -17.424, 33.967]
  MoveL 116 to (362.05, 170.22, 298.54) mm, rotated rx -178.1 ry -46.22 rz 172.02 deg; joints [72.844, 12.364, -28.925, -29.313, -17.576, 34.558]
  MoveL 117 to (361.25, 173.01, 298.54) mm, rotated rx -178.1 ry -46.22 rz 172.02 deg; joints [72.582, 12.558, -28.877, -29.739, -17.731, 35.138]
  MoveL 118 to (360.46, 175.8, 298.54) mm, rotated rx -178.1 ry -46.22 rz 172.02 deg; joints [72.321, 12.751, -28.829, -30.155, -17.887, 35.707]
  MoveL 119 to (359.72, 178.6, 298.54) mm, rotated rx -178.1 ry -46.22 rz 172.02 deg; joints [72.058, 12.939, -28.781, -30.567, -18.045, 36.273]
  MoveL 120 to (359.67, 183.42, 298.54) mm, rotated rx -178.1 ry -46.22 rz 172.02 deg; joints [71.569, 13.127, -28.732, -31.375, -18.307, 37.371]
  MoveL 121 to (361.29, 187.97, 298.54) mm, rotated rx -178.1 ry -46.22 rz 172.02 deg; joints [71.052, 13.118, -28.735, -32.287, -18.544, 38.594]
  MoveL 122 to (364.14, 191.87, 298.54) mm, rotated rx -178.1 ry -46.22 rz 172.02 deg; joints [70.555, 12.947, -28.779, -33.203, -18.742, 39.813]
  MoveL 123 to (367.38, 194.45, 298.54) mm, rotated rx -178.1 ry -46.22 rz 172.02 deg; joints [70.177, 12.682, -28.846, -33.941, -18.87, 40.786]
  MoveL 124 to (371.35, 195.69, 298.54) mm, rotated rx -178.1 ry -46.22 rz 172.02 deg; joints [69.904, 12.281, -28.945, -34.549, -18.922, 41.568]
  MoveL 125 to (375.51, 196.25, 298.54) mm, rotated rx -178.1 ry -46.22 rz 172.02 deg; joints [69.691, 11.83, -29.053, -35.072, -18.94, 42.23]
  MoveL 126 to (379.7, 196.59, 298.54) mm, rotated rx -178.1 ry -46.22 rz 172.02 deg; joints [69.496, 11.367, -29.16, -35.561, -18.951, 42.847]
  MoveL 127 to (383.89, 196.76, 298.54) mm, rotated rx -178.1 ry -46.22 rz 172.02 deg; joints [69.316, 10.896, -29.264, -36.022, -18.959, 43.427]
  MoveL 128 to (388.08, 196.81, 298.54) mm, rotated rx -178.1 ry -46.22 rz 172.02 deg; joints [69.146, 10.421, -29.365, -36.461, -18.965, 43.98]
  MoveL 129 to (392.26, 196.77, 298.54) mm, rotated rx -178.1 ry -46.22 rz 172.02 deg; joints [68.981, 9.941, -29.462, -36.884, -18.973, 44.512]
  MoveL 130 to (400.87, 196.55, 298.54) mm, rotated rx -178.1 ry -46.22 rz 172.02 deg; joints [68.652, 8.948, -29.65, -37.713, -18.997, 45.561]
  MoveL 131 to (409.47, 196.27, 298.54) mm, rotated rx -178.1 ry -46.22 rz 172.02 deg; joints [68.318, 7.95, -29.819, -38.512, -19.043, 46.581]
  MoveL 132 to (418.01, 196.76, 298.54) mm, rotated rx -178.1 ry -46.22 rz 172.02 deg; joints [67.892, 6.991, -29.962, -39.39, -19.164, 47.735]
  MoveL 133 to (426.61, 198.78, 298.54) mm, rotated rx -178.1 ry -46.22 rz 172.02 deg; joints [67.279, 6.099, -30.08, -40.462, -19.414, 49.195]
  MoveL 134 to (431.83, 199.88, 298.54) mm, rotated rx -178.1 ry -46.22 rz 172.02 deg; joints [66.913, 5.552, -30.144, -41.074, -19.573, 50.04]
  MoveL 135 to (435.95, 200.4, 298.54) mm, rotated rx -178.1 ry -46.22 rz 172.02 deg; joints [66.657, 5.103, -30.192, -41.501, -19.682, 50.629]
  MoveL 136 to (439.13, 200.6, 298.54) mm, rotated rx -178.1 ry -46.22 rz 172.02 deg; joints [66.48, 4.747, -30.227, -41.796, -19.758, 51.037]
  MoveL 137 to (441.87, 200.65, 298.54) mm, rotated rx -178.1 ry -46.22 rz 172.02 deg; joints [66.34, 4.433, -30.256, -42.03, -19.817, 51.361]
  MoveL 138 to (444.73, 200.65, 298.54) mm, rotated rx -178.1 ry -46.22 rz 172.02 deg; joints [66.197, 4.103, -30.285, -42.264, -19.878, 51.686]
  MoveL 139 to (447.51, 200.65, 298.54) mm, rotated rx -178.1 ry -46.22 rz 172.02 deg; joints [66.058, 3.782, -30.31, -42.487, -19.941, 51.998]
  MoveL 140 to (451.09, 200.65, 298.54) mm, rotated rx -178.1 ry -46.22 rz 172.02 deg; joints [65.875, 3.368, -30.34, -42.769, -20.025, 52.396]
  MoveL 141 to (455.37, 200.65, 298.54) mm, rotated rx -178.1 ry -46.22 rz 172.02 deg; joints [65.653, 2.871, -30.372, -43.098, -20.133, 52.867]
  MoveL 142 to (459.88, 200.65, 298.54) mm, rotated rx -178.1 ry -46.22 rz 172.02 deg; joints [65.416, 2.348, -30.399, -43.435, -20.253, 53.353]
  Establecer velocidad (1000.0 mm/s)
  MoveL 143 to (459.88, 200.65, 298.54) mm, rotated rx -178.1 ry -46.22 rz 172.02 deg; joints [65.416, 2.348, -30.399, -43.435, -20.253, 53.353]
  MoveL 144 to (479.49, 200.65, 396.6) mm, rotated rx -178.1 ry -46.22 rz 172.02 deg; joints [64.329, -4.285, -16.18, -27.823, -32.517, 36.529]

